(* IEC 61131-3 sources: daoli-st-library/DL_Device (part 42) *)

(* ---- FB_DL_PumpCavitationGuard.st ---- *)
(*==============================================================================
 * 组件名称 (Component)  : FB_DL_PumpCavitationGuard
 * 所属子库 (Sublibrary) : DL_Device
 * 当前版本 (Version)    : 1.0.1
 * 兼容性   (Platform)   : CODESYS 3.5 / TwinCAT 3 / 汇川 InoProShop / Schneider
 *                         Machine Expert；纯 IEC 61131-3（第 3 版）语法，
 *                         仅依赖 Standard.library（R_TRIG / TON）
 * 组件分类 (Category)   : 功能块（FUNCTION_BLOCK）· 设备本体退化诊断 · 泵汽蚀
 * 功能描述 (Function)   : 泵汽蚀的在线判据与**降速请求**。三判据并发：
 *                         (a) 流量偏低（低于额定的比例）；(b) 扬程跌落（低于额定的
 *                         跌幅）；(c) 振动超限**或**电流波动超限。三者同拍成立并
 *                         持续 tConfirm 才升级为锁存故障；单条成立只到「嫌疑」。
 * 降速语义 (Derate)     : 本件**不直接给变频器频率**，只输出 `fDerateRatio`
 *                         （1.0 = 不降）与 `bDerateRequest`。执行归上层
 *                         `FB_DL_RateLimiter` / `FB_DL_VfdGeneric`——诊断件一旦
 *                         自己写频率，就会与工艺主控的速率限制打架，且无法在
 *                         不同变频器之间移植。
 *                         每次确认汽蚀事件比率递减一步（下限 0.3），**只减不自动
 *                         增**：回升由上层斜坡完成，避免本件与上层同时调节同
 *                         一个量（双写冲突）。
 * 边界声明 (Limits)     : ① **不做 NPSH 计算**：需介质饱和蒸汽压与吸入侧压力，
 *                         属选型设计而非在线判据；② 振动阈值默认取 ISO 10816
 *                         C 区边界 4.5 mm/s（**公知阈值，引脚可改**），头注释
 *                         注明出处与「仅参考」定位；③ 本件**不声称**符合
 *                         ISO 10816 认证，阈值只是工程默认值；④ 停泵（bRunning
 *                         为 FALSE）时全部判据抑制，不产生任何降速请求。
 * 段序 (Cycle order)   : 段 1 默认值与单拍预清零 → 段 2 首扫初始化 →
 *                         段 3 参数闸门与输入域检查 → 段 4 定时器与边沿无条件刷新 →
 *                         段 5 判据计算 → 段 6 复位通道与故障锁存（**CASE 前置，
 *                         不做状态变量赋值**）→ 段 7 监视相位机 → 段 8 降速执行与
 *                         事件锁存 → 段 9 健康仲裁、出口钳位与保持重写 → 段 10 码位链。
 * 拍间依赖 (Cycle dep)  : 确认定时器在段 4 调用，而其 IN 里的「三判据同拍」在段 5
 *                         才算出，故定时器读到的是**上一拍照**的判据值（一拍滞后）。
 *                         对 3 秒量级的确认判据无实质影响，换来的是「所有定时器
 *                         实例都在同一段无条件调用」这一更强的纪律；此处显式登记，
 *                         避免后人误以为是笔误。
 * 定时器清单 (R40)      : 实例名 / IN 表达式 / 断输入拍标志 / 自清位置
 *                         fbConfirmWatch / 三判据同拍 AND 状态为嫌疑 AND
 *                                        NOT _bConfirmBreak / _bConfirmBreak
 *                                        （进/出嫌疑态与复位时置位）
 *                         fbRippleWatch  / 泵运行 AND NOT _bRippleBreak
 *                                        / _bRippleBreak（窗满后置位重启）
 *                         fbHoldOffWatch / 状态为降速 AND NOT _bHoldBreak
 *                                        / _bHoldBreak（进/出降速态置位）
 *                         三个实例全部在段 4 无条件调用，断输入拍一律在调用后自清。
 * 单拍标志清单 (R25)    : `_bResetPulse` 预清段 1 / 置位段 6 / 消费段 6；
 *                         `_bDerateStep`（降速单拍）预清段 1 / 置位段 8 / 消费段 8；
 *                         `_bConfirmEvent` 预清段 1 / 置位段 7 / 消费段 8；
 *                         三个断输入标志就地置位、段 4 调用后自清。
 * 保持位清单 (R27)      : `bDerateRequest` 与 `fDerateRatio`、`bCavitation`、
 *                         `nEventCount` 四个保持量，全部由段 9 每拍重写出口；
 *                         降速请求在 eDerate 与抑制窗内**保持为 TRUE**，不靠
 *                         进入那一拍的脉冲（R27 的典型场景）。
 * 三元一致表 (R35)      : 量 / 守卫封顶 / 判据运算符
 *                         fFlowLowRatio   / 钳到 0.2~0.95 / 判据用 <
 *                         fHeadDropRatio  / 钳到 0.05~0.5 / 判据用（1 减比值）>
 *                         fVibLimit       / 钳到 1~20     / 判据用比值 > 1，急停用 > 2
 *                         振动比值输出上限 / 钳到 5.0     / 必须高于急停倍率 2（R35 同向）
 *                         fDerateStep     / 钳到 0.02~0.3 / 递减后与 0.3 取大
 * 验收向量 (Acceptance) :
 *   V1 单判据：流量 0.5 倍额定（其余判据不成立）→ eSuspect + 0164，**不锁存**
 *   V2 三判据：三判据同拍持续 3 s → eConfirm → eDerate、0326、比率每次 −0.10
 *      （下限 0.3）
 *   V3（V-C 跨段 R40）：tConfirm 定时器在 eSuspect 与 eMonitor 来回时必须断输入，
 *      否则三次 1 s 的孤立嫌疑会被误判成「持续 3 s」
 *   V4（V-D 恢复）：bReset 后 fDerateRatio **不得**直接回 1.0（R41），且必须夹进
 *      0.3~1.0（R43）
 *   V5（V-A 域外）：fFlowNominal 为 0 → 0328 锁存，fFlowRatio 输出 0（不输出无穷大）
 * 规格偏离 (Deviation)  :
 *   ① 规格 V1 给的是「流量 0.5 倍额定、扬程 0.8 倍额定、振动 2.0、电流平稳 →
 *      只有流量判据」。按默认 fHeadDropRatio 为 0.15 计算，扬程 0.8 倍额定的跌幅
 *      为 20%，**会同时触发扬程判据**。本件按判据定义实现（跌幅 > 15% 即成立），
 *      复现 V1 需把 fHeadDropRatio 调到 ≥0.25；此处不改判据语义以迁就向量。
 *   ② 规格未给「电流波动率」的确切口径。本件取滑动窗内「(最大 − 最小) ÷ 平均」
 *      作为波动率，窗长 tRippleWindow，窗满即出值并重启窗；该口径与现场常见的
 *      「电流摆动幅度百分比」一致，且不依赖频谱。
 *   ③ 规格要求 bReset 后比率不直接回 1.0。本件在 bReset 且三判据全部消失时让
 *      比率**回升一步**（不直接回 1.0），其余恢复速率仍交上层斜坡；这是「不得
 *      重头恢复」与「不能让比率永久卡死」之间的折中，已在此登记。
 *   ④ 参数非法（额定值非正、阈值倒置）统一用 0328，未分更细码位（本轮未分配）。
 * 开源溯源 (Origin)     : 来源标签 namur-ne107 / lbp-basic-process / pump-diag。
 *                         原创 clean-room 实现。**仅借鉴**：① NAMUR NE107（公开
 *                         推荐规范）的健康分级语义；② LBP（Library of Basic
 *                         Process）公开文档所呈现的「命令—监视—判定」三段式
 *                         分层惯例，作为本件「判据—定级—降速请求」的组织参照。
 *                         汽蚀三判据（流量低 / 扬程跌 / 振动或电流波动）属泵
 *                         行业公开的通行定性认识；ISO 10816 的 4.5 mm/s 为公知
 *                         阈值。本件未复制任何源码行、未沿用其命名体系，窗口
 *                         口径、状态机、宽限与降速规则、全部码位 100% 本库独立
 *                         设计，无许可证传染风险。
 * 修订历史 (Revision)   :
 *   2026-11-15  v1.0.0  首版入库（R13 · 泳道 A · 泵汽蚀判据与降速请求）
 *   2026-11-16  v1.0.1  终审修复五处：① `_bHoldActive` 由「窗满那一拍」改为
 *                       「整个降速相」——原实现下 0165 仅在抑制窗到期瞬间可见、
 *                       判据在窗内并未被真正抑制；② 流量/扬程比值改用**原始
 *                       额定值的域**做门（原实现拿兜底值 1.0 当分母，额定为 0
 *                       时输出的是伪比值而非 0，违 V5）；③ 汽蚀确认补写
 *                       `_uErrFault := 16#0003_0326`（原实现 bError 为真而
 *                       uErrorId 恒 0，违 R21 一致性）；④ 急停级 0327 加
 *                       bRunning/bEnable 门（停泵时邻近设备振动不得拉锁存）；
 *                       ⑤ 停泵清 `_fRipple`，防停泵前旧波动率跨停机存活到
 *                       重启后的首个取样窗。
 *============================================================================*)

(*-----------------------------------------------------------------------------
 * 枚举: E_DL_CavitationState（归属本功能块，同文件发布）
 * 含义: 汽蚀监视相位。6 个成员在段 6 各有唯一标签，ELSE 只接脏值。
 *-----------------------------------------------------------------------------*)
TYPE E_DL_CavitationState :
(
    eIdle    := 0,     // 待机：未使能或停泵 / Idle, disabled or the pump is stopped
    eMonitor := 10,    // 监视：泵运行，判据全部不成立 / Monitoring, no criterion active
    eSuspect := 20,    // 嫌疑：单判据成立，未确认 / Suspect, one criterion active
    eConfirm := 30,    // 确认：三判据同拍且持续满足 / Confirm, all three held long enough
    eDerate  := 40,    // 降速：已请求降速，处于抑制窗 / Derate, request held during the hold-off
    eFault   := 99     // 故障：参数非法或振动急停级，锁存 / Fault, latched
);
END_TYPE

FUNCTION_BLOCK FB_DL_PumpCavitationGuard
VAR_INPUT
    bEnable             : BOOL;                      // 使能 [-] / Enable
    bReset              : BOOL;                      // 复位锁存，上升沿有效 [-] / Rising edge resets the latch
    bRunning            : BOOL;                      // 泵运行中，停泵时全部判据抑制 [-] / Pump running, criteria suppressed when stopped
    fFlow               : REAL;                      // 实测流量 [m³/h]，范围 0~100000 / Measured flow
    fHead               : REAL;                      // 实测扬程 [m]，范围 0~1000 / Measured head
    fVibration          : REAL;                      // 振动速度有效值 [mm/s]，范围 0~50 / Vibration RMS velocity
    fCurrent            : REAL;                      // 电机电流 [A]，范围 0~10000 / Motor current
    fFlowNominal        : REAL;                      // 额定流量 [m³/h]，域大于 0 / Nominal flow, must exceed zero
    fHeadNominal        : REAL;                      // 额定扬程 [m]，域大于 0 / Nominal head, must exceed zero
    fFlowLowRatio       : REAL := 0.60;              // 流量低于额定的比例 [-]，范围 0.2~0.95 / Low-flow ratio
    fHeadDropRatio      : REAL := 0.15;              // 扬程跌落比例 [-]，范围 0.05~0.5 / Head-drop ratio
    fVibLimit           : REAL := 4.5;               // 振动上限 [mm/s]，ISO 10816 C 区边界，范围 1~20 / Vibration limit
    fCurrentRippleLimit : REAL := 0.15;              // 电流波动率上限 [-]，范围 0.02~0.5 / Current ripple limit
    tRippleWindow       : TIME := T#2S;              // 电流波动统计窗 [毫秒]，范围 0.5~30 s / Ripple window
    tConfirm            : TIME := T#3S;              // 三判据同拍持续判据 [毫秒]，范围 0.5~30 s / Confirmation time
    tHoldOff            : TIME := T#30S;             // 降速后抑制判据时长 [毫秒]，范围 5 s~10 min / Hold-off after a derate
    fDerateStep         : REAL := 0.10;              // 每次降速步长 [-]，范围 0.02~0.3 / Derate step
END_VAR
VAR_OUTPUT
    eHealth             : E_DL_Ne107Status;          // NE107 健康态（引用自 I_DL_DeviceHealth）[-] / NE107 health
    uDiagCode           : UDINT;                     // 当前诊断码，0=无码 [代码] / Active diagnostic code
    uErrorId            : UDINT;                     // 末次故障码，仅故障级 [代码] / Last fault code
    bError              : BOOL;                      // 故障锁存 [-] / Fault latched
    bCavitation         : BOOL;                      // 汽蚀确认（三判据同拍成立，锁存）[-] / Cavitation confirmed, latched
    bDerateRequest      : BOOL;                      // 降速请求（保持语义）[-] / Derate request, held
    fDerateRatio        : REAL;                      // 降速比例 [-]，范围 0.3~1.0，1.0=不降 / Derate ratio
    fFlowRatio          : REAL;                      // 实测/额定流量比值 [-]，钳 0~2 / Flow ratio
    fHeadRatio          : REAL;                      // 实测/额定扬程比值 [-]，钳 0~2 / Head ratio
    fVibRatio           : REAL;                      // 振动/上限比值 [-] / Vibration ratio
    nEventCount         : UDINT;                     // 汽蚀事件累计 [次]，锁存 / Event counter
    fRippleMeas         : REAL;                      // 窗内电流波动率实测值 [-] / Measured ripple
END_VAR
VAR
    fbTrigReset     : R_TRIG;                        // 复位沿检测，段 4 无条件刷新 [-] / Reset edge detector
    fbConfirmWatch  : TON;                           // 三判据持续计时，段 4 刷新 [毫秒] / Confirmation timer
    fbRippleWatch   : TON;                           // 电流波动统计窗，段 4 刷新 [毫秒] / Ripple window timer
    fbHoldOffWatch  : TON;                           // 降速后抑制窗，段 4 刷新 [毫秒] / Hold-off timer
    _eState         : E_DL_CavitationState := E_DL_CavitationState.eIdle; // 当前相位 [-] / Current phase
    _bInit          : BOOL := FALSE;                 // 首扫标志，初值 FALSE [-] / First-scan flag
    _bFaultLatch    : BOOL;                          // 故障锁存，仅复位清 [-] / Fault latch
    _uErrFault      : UDINT;                         // 首出故障码 [代码] / First-out fault code
    _uDiagCode      : UDINT;                         // 当前诊断码（单一链产出）[代码] / Active diagnostic code
    _bResetPulse    : BOOL;                          // 复位单拍 [-] / One-shot reset
    _bParamBad      : BOOL;                          // 参数非法标志 [-] / Illegal parameter flag
    _bConfirmBreak  : BOOL;                          // 确认定时器断输入一拍 [-] / Confirmation timer break
    _bRippleBreak   : BOOL;                          // 波动窗断输入一拍 [-] / Ripple window break
    _bHoldBreak     : BOOL;                          // 抑制窗断输入一拍 [-] / Hold-off break
    _fFlowNomUse    : REAL := 1.0;                   // 生效额定流量 [m³/h] / Effective nominal flow
    _fHeadNomUse    : REAL := 1.0;                   // 生效额定扬程 [m] / Effective nominal head
    _fFlowLowUse    : REAL := 0.60;                  // 生效流量比例 [-] / Effective low-flow ratio
    _fHeadDropUse   : REAL := 0.15;                  // 生效扬程跌幅 [-] / Effective head-drop ratio
    _fVibUse        : REAL := 4.5;                   // 生效振动上限 [mm/s] / Effective vibration limit
    _fRippleLimUse  : REAL := 0.15;                  // 生效波动率上限 [-] / Effective ripple limit
    _fStepUse       : REAL := 0.10;                  // 生效降速步长 [-] / Effective derate step
    _tRippleUse     : TIME := T#2S;                  // 生效波动窗 [毫秒] / Effective ripple window
    _tConfirmUse    : TIME := T#3S;                  // 生效确认时长 [毫秒] / Effective confirmation time
    _tHoldUse       : TIME := T#30S;                 // 生效抑制窗 [毫秒] / Effective hold-off
    _diMs           : DINT;                          // 时间换算中间量 [毫秒] / Time conversion working value
    _fFlowRatio     : REAL;                          // 流量比值 [-]，钳 0~2 / Flow ratio
    _fHeadRatio     : REAL;                          // 扬程比值 [-]，钳 0~2 / Head ratio
    _fVibRatio      : REAL;                          // 振动比值 [-] / Vibration ratio
    _bCritFlow      : BOOL;                          // 流量判据 [-] / Flow criterion
    _bCritHead      : BOOL;                          // 扬程判据 [-] / Head criterion
    _bCritVib       : BOOL;                          // 振动判据 [-] / Vibration criterion
    _bCritRipple    : BOOL;                          // 电流波动判据 [-] / Ripple criterion
    _bCritVibGroup  : BOOL;                          // 振动或波动（第三判据）[-] / Vibration or ripple, the third criterion
    _bAllThree      : BOOL;                          // 三判据同拍成立 [-] / All three criteria in one scan
    _bAnyCrit       : BOOL;                          // 任一判据成立 [-] / Any criterion active
    _bVibEmergency  : BOOL;                          // 振动超上限两倍（急停级）[-] / Vibration above twice the limit
    _fCurrMin       : REAL;                          // 窗内电流最小值 [A] / Minimum current in the window
    _fCurrMax       : REAL;                          // 窗内电流最大值 [A] / Maximum current in the window
    _fCurrSum       : REAL;                          // 窗内电流累加 [A] / Current sum in the window
    _nCurrCount     : UDINT;                         // 窗内电流样本数 [个] / Current sample count
    _fRipple        : REAL;                          // 窗内波动率实测值 [-] / Measured ripple
    _bHoldActive    : BOOL;                          // 抑制窗生效中 [-] / Hold-off active
    _bDerateStep    : BOOL;                          // 本次确认需降一步 [-] / Step down this scan
    _bConfirmEvent  : BOOL;                          // 本拍确认事件 [-] / Confirmation event this scan
    _bCavLatch      : BOOL;                          // 汽蚀锁存 [-] / Cavitation latch
    _fDerateRatio   : REAL := 1.0;                   // 保持的降速比例 [-] / Held derate ratio
    _bDerateHeld    : BOOL;                          // 保持的降速请求 [-] / Held derate request
    _uEventCount    : UDINT;                         // 保持的事件计数 [次] / Held event counter
    _eHealthInt     : E_DL_Ne107Status := E_DL_Ne107Status.eUnknown; // 健康态内部量 [-] / Internal health state
END_VAR
VAR CONSTANT
    DL_VAL_LIM      : REAL := 1.0E6;                 // 有限性判定绝对值上限 [-] / Finiteness limit
    DL_EPS          : REAL := 1.0E-6;                // 浮点比较容差 [-] / Float comparison tolerance
    DL_RATIO_MAX    : REAL := 2.0;                   // 流量扬程比值上限 [-]，防噪声放大 / Flow and head ratio ceiling
    DL_VIB_RATIO_MAX: REAL := 5.0;                   // 振动比值上限 [-]，须高于急停倍率 2 倍（R35 同向） / Vibration ratio ceiling
    DL_VIB_EMERG    : REAL := 2.0;                   // 振动急停级倍率 [-] / Emergency vibration multiplier
    DL_DERATE_MIN   : REAL := 0.3;                   // 降速比例下限 [-] / Lower derate bound
    DL_DERATE_MAX   : REAL := 1.0;                   // 降速比例上限 [-] / Upper derate bound
    DL_RIPPLE_MIN_MS: DINT := 500;                   // 波动窗下限 [毫秒] / Minimum ripple window
    DL_RIPPLE_MAX_MS: DINT := 30000;                 // 波动窗上限 [毫秒] / Maximum ripple window
    DL_CONFIRM_MIN  : DINT := 500;                   // 确认时长下限 [毫秒] / Minimum confirmation
    DL_CONFIRM_MAX  : DINT := 30000;                 // 确认时长上限 [毫秒] / Maximum confirmation
    DL_HOLD_MIN     : DINT := 5000;                  // 抑制窗下限 [毫秒] / Minimum hold-off
    DL_HOLD_MAX     : DINT := 600000;                // 抑制窗上限 [毫秒] / Maximum hold-off
END_VAR

(*------------------------------------------------------------------------------
 * 段 1｜确定性默认值与单拍标志预清零（R25 第一律）
 *      Deterministic defaults and one-shot flags pre-cleared
 *-----------------------------------------------------------------------------*)
_bResetPulse   := FALSE;                              // 复位单拍预清零（Reset pre-cleared）
_bParamBad     := FALSE;                              // 参数非法预清零（Illegal parameter pre-cleared）
_bDerateStep   := FALSE;                              // 降速单拍预清零（Derate step pre-cleared）
_bConfirmEvent := FALSE;                              // 确认事件预清零（Confirmation event pre-cleared）
_bCritFlow     := FALSE;                              // 流量判据预清零（Flow criterion pre-cleared）
_bCritHead     := FALSE;                              // 扬程判据预清零（Head criterion pre-cleared）
_bCritVib      := FALSE;                              // 振动判据预清零（Vibration criterion pre-cleared）
_bCritRipple   := FALSE;                              // 波动判据预清零（Ripple criterion pre-cleared）
_bVibEmergency := FALSE;                              // 振动急停预清零（Emergency pre-cleared）

(*------------------------------------------------------------------------------
 * 段 2｜首扫初始化（R19：bInit 初值 FALSE，判据取非；首拍只装基准）
 *      First-scan initialisation, baseline only
 *-----------------------------------------------------------------------------*)
IF NOT _bInit THEN
    _eState       := E_DL_CavitationState.eIdle;      // 相位待机（Phase idle）
    _bFaultLatch  := FALSE;                           // 故障锁存清零（Latch cleared）
    _uErrFault    := 16#0000_0000;                    // 首出码清零（First-out code cleared）
    _bCavLatch    := FALSE;                           // 汽蚀锁存清零（Cavitation latch cleared）
    _fDerateRatio := DL_DERATE_MAX;                   // 冷启动比率 1.0，落在有效域内（Cold start at 1.0）
    _bDerateHeld  := FALSE;                           // 降速请求清零（Derate request cleared）
    _uEventCount  := 0;                               // 事件计数清零（Event counter cleared）
    _fRipple      := 0.0;                             // 波动率初值 0（Ripple starts at zero）
    _fCurrMin     := DL_VAL_LIM;                      // 最小值先置上界（Minimum preset to the ceiling）
    _fCurrMax     := 0.0;                             // 最大值先置 0（Maximum preset to zero）
    _fCurrSum     := 0.0;                             // 电流累加清零（Current sum cleared）
    _nCurrCount   := 0;                               // 样本数清零（Sample count cleared）
    _fFlowNomUse  := 1.0;                             // 额定流量兜底（Nominal flow fallback）
    _fHeadNomUse  := 1.0;                             // 额定扬程兜底（Nominal head fallback）
    _bInit        := TRUE;                            // 首扫只做一次（First scan runs once）
END_IF

(*------------------------------------------------------------------------------
 * 段 3｜参数闸门与输入域检查（额定值非正或阈值倒置属故障级）
 *      Parameter gate: non-positive nominals or inverted thresholds latch a fault
 *-----------------------------------------------------------------------------*)
IF (fFlowNominal <= DL_EPS) OR (fHeadNominal <= DL_EPS) OR (fVibLimit <= DL_EPS) THEN
    _bParamBad := TRUE;                               // 额定值或振动上限非正（Non-positive nominals）
END_IF
IF (fFlowLowRatio <= 0.0) OR (fFlowLowRatio >= 1.0) OR (fHeadDropRatio <= 0.0) OR (fHeadDropRatio >= 1.0) THEN
    _bParamBad := TRUE;                               // 比例阈值倒置（Inverted ratios）
END_IF
IF (fCurrentRippleLimit <= 0.0) OR (fDerateStep <= 0.0) OR (fDerateStep > 0.5) THEN
    _bParamBad := TRUE;                               // 波动限或步长非法（Illegal ripple limit or step）
END_IF

IF fFlowNominal > DL_EPS THEN
    _fFlowNomUse := fFlowNominal;                     // 额定流量直通（Nominal flow passed through）
ELSE
    _fFlowNomUse := 1.0;                              // 非正：兜底为 1，防除零（Fallback avoids a zero divisor）
END_IF
IF fHeadNominal > DL_EPS THEN
    _fHeadNomUse := fHeadNominal;                     // 额定扬程直通（Nominal head passed through）
ELSE
    _fHeadNomUse := 1.0;                              // 非正：兜底为 1（Fallback）
END_IF

_fFlowLowUse   := LIMIT(0.2, fFlowLowRatio, 0.95);    // 流量比例钳进 0.2~0.95（Clamped）
_fHeadDropUse  := LIMIT(0.05, fHeadDropRatio, 0.5);   // 跌幅比例钳进 0.05~0.5（Clamped）
_fVibUse       := LIMIT(1.0, fVibLimit, 20.0);        // 振动上限钳进 1~20 mm/s（Clamped）
_fRippleLimUse := LIMIT(0.02, fCurrentRippleLimit, 0.5); // 波动限钳进 0.02~0.5（Clamped）
_fStepUse      := LIMIT(0.02, fDerateStep, 0.3);      // 降速步长钳进 0.02~0.3（Clamped）

_diMs         := LIMIT(DL_RIPPLE_MIN_MS, TIME_TO_DINT(tRippleWindow), DL_RIPPLE_MAX_MS); // 波动窗钳位（Clamped）
_tRippleUse   := DINT_TO_TIME(_diMs);                 // 生效波动窗（Effective ripple window）
_diMs         := LIMIT(DL_CONFIRM_MIN, TIME_TO_DINT(tConfirm), DL_CONFIRM_MAX); // 确认时长钳位（Clamped）
_tConfirmUse  := DINT_TO_TIME(_diMs);                 // 生效确认时长（Effective confirmation）
_diMs         := LIMIT(DL_HOLD_MIN, TIME_TO_DINT(tHoldOff), DL_HOLD_MAX); // 抑制窗钳位（Clamped）
_tHoldUse     := DINT_TO_TIME(_diMs);                 // 生效抑制窗（Effective hold-off）

(*------------------------------------------------------------------------------
 * 段 4｜定时器与边沿实例无条件刷新（红线：实例一律在 CASE 之外每拍必调）
 *      Timers and edge detectors refreshed unconditionally outside the CASE
 *-----------------------------------------------------------------------------*)
fbTrigReset(CLK := bReset);                           // 复位沿刷新（Reset edge refreshed）

fbConfirmWatch(IN := _bAllThree AND (_eState = E_DL_CavitationState.eSuspect) AND (NOT _bConfirmBreak), PT := _tConfirmUse); // 三判据持续计时
_bConfirmBreak := FALSE;                              // 断输入拍在调用后自清（Break self-cleared）

fbRippleWatch(IN := bRunning AND (NOT _bRippleBreak), PT := _tRippleUse); // 波动统计窗
_bRippleBreak := FALSE;                               // 断输入拍在调用后自清（Break self-cleared）

fbHoldOffWatch(IN := (_eState = E_DL_CavitationState.eDerate) AND (NOT _bHoldBreak), PT := _tHoldUse); // 抑制窗计时
_bHoldBreak := FALSE;                                 // 断输入拍在调用后自清（Break self-cleared）
_bHoldActive := (_eState = E_DL_CavitationState.eDerate) OR fbHoldOffWatch.Q; // 抑制生效 = 整个降速相（不是窗满那一拍）

(*------------------------------------------------------------------------------
 * 段 5｜判据计算（比值前置守卫，绝不输出无穷大；V5）
 *      Criteria, ratios guarded against division by zero
 *-----------------------------------------------------------------------------*)
(* 比值口径：额定值非正时**输出 0**，绝不拿兜底值 1.0 去算伪比值（V5 明确要求） *)
IF fFlowNominal > DL_EPS THEN
    _fFlowRatio := LIMIT(0.0, fFlow / _fFlowNomUse, DL_RATIO_MAX); // 流量比值，钳 0~2（Clamped）
ELSE
    _fFlowRatio := 0.0;                               // 额定流量非法：输出 0，不给伪比值（Never a pseudo ratio）
END_IF
IF fHeadNominal > DL_EPS THEN
    _fHeadRatio := LIMIT(0.0, fHead / _fHeadNomUse, DL_RATIO_MAX); // 扬程比值，钳 0~2（Clamped）
ELSE
    _fHeadRatio := 0.0;                               // 额定扬程非法：输出 0（Never a pseudo ratio）
END_IF
IF _fVibUse > DL_EPS THEN
    _fVibRatio := LIMIT(0.0, fVibration / _fVibUse, DL_VIB_RATIO_MAX); // 振动比值，上限须容得下急停倍率（Clamped）
ELSE
    _fVibRatio := 0.0;                                // 分母不可用：输出 0（Never infinity）
END_IF

(* 三判据：停泵或抑制窗内一律不成立（Suppressed when stopped or within the hold-off） *)
IF bRunning AND bEnable AND (NOT _bHoldActive) THEN
    _bCritFlow   := _fFlowRatio < _fFlowLowUse;                       // 流量偏低（Low flow）
    _bCritHead   := _fHeadRatio < (1.0 - _fHeadDropUse);              // 扬程跌落（Head drop）
    _bCritVib    := _fVibRatio > 1.0;                                 // 振动超限（Vibration above limit）
    _bCritRipple := _fRipple > _fRippleLimUse;                        // 电流波动超限（Ripple above limit）
END_IF
_bCritVibGroup := _bCritVib OR _bCritRipple;                          // 第三判据：振动或波动（Third criterion）
_bAllThree     := _bCritFlow AND _bCritHead AND _bCritVibGroup;       // 三判据同拍（All three in one scan）
_bAnyCrit      := _bCritFlow OR _bCritHead OR _bCritVibGroup;         // 任一判据（Any criterion）
(* 急停级：仅在泵运行且使能时成立。停泵时邻近设备振动/传感器卡值不得把本件拉进锁存，
 * 与「bRunning 为 FALSE 时全部判据抑制」同一条纪律；降速抑制窗内仍照判（等级高于判据） *)
IF bRunning AND bEnable AND (_fVibRatio > DL_VIB_EMERG) THEN
    _bVibEmergency := TRUE;                                           // 振动超两倍上限（Emergency level）
END_IF

(* 电流波动统计：窗满出一值并重启窗（Window closes, one value produced, window restarts） *)
IF bRunning THEN
    IF fCurrent < _fCurrMin THEN
        _fCurrMin := fCurrent;                        // 更新最小（Update the minimum）
    END_IF
    IF fCurrent > _fCurrMax THEN
        _fCurrMax := fCurrent;                        // 更新最大（Update the maximum）
    END_IF
    _fCurrSum := _fCurrSum + fCurrent;                // 累加（Accumulate）
    IF _nCurrCount < 16#FFFF_FFFF THEN
        _nCurrCount := _nCurrCount + 1;               // 计数防上溢（Guard the counter）
    END_IF
    IF fbRippleWatch.Q THEN
        IF _nCurrCount > 0 THEN
            IF (_fCurrSum / UDINT_TO_REAL(_nCurrCount)) > DL_EPS THEN
                _fRipple := (_fCurrMax - _fCurrMin) / (_fCurrSum / UDINT_TO_REAL(_nCurrCount)); // 波动率，分母已守卫
            ELSE
                _fRipple := 0.0;                      // 平均近零：不判波动（No meaningful ripple）
            END_IF
        END_IF
        _fCurrMin   := DL_VAL_LIM;                    // 窗重启：最小值复位（Window restarted）
        _fCurrMax   := 0.0;                           // 窗重启：最大值复位（Window restarted）
        _fCurrSum   := 0.0;                           // 窗重启：累加清零（Window restarted）
        _nCurrCount := 0;                             // 窗重启：计数清零（Window restarted）
        _bRippleBreak := TRUE;                        // 断输入一拍后重新计时（One-scan break restarts the timer）
    END_IF
ELSE
    _fCurrMin   := DL_VAL_LIM;                        // 停泵清零（Cleared while stopped）
    _fCurrMax   := 0.0;                               // 停泵清零（Cleared while stopped）
    _fCurrSum   := 0.0;                               // 停泵清零（Cleared while stopped）
    _nCurrCount := 0;                                 // 停泵清零（Cleared while stopped）
    _fRipple    := 0.0;                               // 停泵清实测值，防停泵前旧值跨停机存活（Stale ripple must not survive a stop）
END_IF

(*------------------------------------------------------------------------------
 * 段 6｜复位通道 + 故障锁存（CASE 前置；**不做状态变量赋值**，R39）
 *      Reset channel and fault latching before the CASE, with no state write
 *-----------------------------------------------------------------------------*)
IF fbTrigReset.Q THEN
    _bResetPulse := TRUE;                             // 复位单拍（One-shot reset）
END_IF

IF _bResetPulse THEN
    _bFaultLatch := FALSE;                            // 清故障锁存（Latch cleared）
    _uErrFault   := 16#0000_0000;                     // 清首出码（First-out code cleared）
    _bCavLatch   := FALSE;                            // 清汽蚀锁存（Cavitation latch cleared）
    _bDerateHeld := FALSE;                            // 撤降速请求，交给上层斜坡（Release the request to the upper ramp）
    IF _bAnyCrit THEN
        _fDerateRatio := LIMIT(DL_DERATE_MIN, _fDerateRatio, DL_DERATE_MAX); // 判据仍在：比率保持并夹域（Held while criteria persist）
    ELSE
        _fDerateRatio := LIMIT(DL_DERATE_MIN, _fDerateRatio + _fStepUse, DL_DERATE_MAX); // 判据已消：回升一步，不直接回 1.0（R41）
    END_IF
    _bConfirmBreak := TRUE;                           // 确认计时重启（Confirmation timer restarted）
    _bRippleBreak  := TRUE;                           // 波动窗重启（Ripple window restarted）
    _bHoldBreak    := TRUE;                           // 抑制窗重启（Hold-off restarted）
END_IF

IF _bParamBad AND (NOT _bFaultLatch) THEN
    _uErrFault   := 16#0003_0328;                     // 0328 额定值非正或阈值倒置（Illegal nominals or thresholds）
    _bFaultLatch := TRUE;                             // 锁存（Latched）
END_IF

(*------------------------------------------------------------------------------
 * 段 7｜监视相位机（6 个成员各一标签 + ELSE 兜底）
 *      Monitoring state machine, one label per member plus a trailing fallback
 *-----------------------------------------------------------------------------*)
CASE _eState OF

    E_DL_CavitationState.eIdle: // 待机：起泵后进入监视
        IF _bFaultLatch THEN
            _eState := E_DL_CavitationState.eFault;   // 已锁故障（Already latched）
        ELSIF bEnable AND bRunning THEN
            _bConfirmBreak := TRUE;                   // 确认计时从 0 起算（Confirmation restarts）
            _bRippleBreak  := TRUE;                   // 波动窗从 0 起算（Ripple window restarts）
            _bHoldBreak    := TRUE;                   // 抑制窗从 0 起算（Hold-off restarts）
            _eState := E_DL_CavitationState.eMonitor; // 进监视（Enter monitoring）
        END_IF

    E_DL_CavitationState.eMonitor: // 监视：任一判据即进嫌疑
        IF _bFaultLatch THEN
            _eState := E_DL_CavitationState.eFault;   // 转故障（Enter the fault state）
        ELSIF (NOT bEnable) OR (NOT bRunning) THEN
            _eState := E_DL_CavitationState.eIdle;    // 停泵或掉使能回待机（Stopped or disabled, back to idle）
        ELSIF _bAnyCrit AND (NOT _bHoldActive) THEN
            _bConfirmBreak := TRUE;                   // 进嫌疑：确认计时从 0 起算（R40 段边界断输入）
            _eState := E_DL_CavitationState.eSuspect; // 进嫌疑（Enter suspect）
        END_IF

    E_DL_CavitationState.eSuspect: // 嫌疑：三判据同拍并持续满足才确认
        IF _bFaultLatch THEN
            _eState := E_DL_CavitationState.eFault;   // 转故障（Enter the fault state）
        ELSIF (NOT bEnable) OR (NOT bRunning) THEN
            _eState := E_DL_CavitationState.eIdle;    // 停泵回待机（Stopped, back to idle）
        ELSIF NOT _bAnyCrit THEN
            _bConfirmBreak := TRUE;                   // 判据消失：确认计时断输入（Criterion cleared, timer broken）
            _eState := E_DL_CavitationState.eMonitor; // 回监视（Back to monitoring）
        ELSIF fbConfirmWatch.Q THEN
            _bConfirmEvent := TRUE;                   // 确认事件单拍（Confirmation event）
            _eState := E_DL_CavitationState.eConfirm; // 进确认（Enter confirmation）
        END_IF

    E_DL_CavitationState.eConfirm: // 确认：本拍锁存并请求降速，随后进入降速相
        _bConfirmBreak := TRUE;                       // 确认计时清零（Confirmation cleared）
        _bHoldBreak    := TRUE;                       // 抑制窗从 0 起算（Hold-off restarts）
        _eState := E_DL_CavitationState.eDerate;      // 进降速（Enter derate）
        IF (NOT bEnable) OR (NOT bRunning) THEN
            _eState := E_DL_CavitationState.eIdle;    // 停泵中止（Stopped, abort）
        END_IF

    E_DL_CavitationState.eDerate: // 降速：抑制窗内忽略判据，窗满且判据消失才回监视
        IF _bFaultLatch THEN
            _eState := E_DL_CavitationState.eFault;   // 转故障（Enter the fault state）
        ELSIF (NOT bEnable) OR (NOT bRunning) THEN
            _bHoldBreak := TRUE;                      // 抑制窗中断（Hold-off stopped）
            _eState := E_DL_CavitationState.eIdle;    // 停泵回待机（Stopped, back to idle）
        ELSIF fbHoldOffWatch.Q THEN
            (* 抑制窗内判据被强制为假，故出口条件只看窗满；窗满后判据在
             * eMonitor 重新评估，若仍成立会再次进入嫌疑并再降一步 *)
            _bHoldBreak := TRUE;                      // 抑制窗结束重启（Hold-off finished）
            _bDerateHeld := FALSE;                    // 撤降速请求，交由上层斜坡（Request released to the upper ramp）
            _bConfirmBreak := TRUE;                   // 确认计时重启（Confirmation restarted）
            _eState := E_DL_CavitationState.eMonitor; // 回监视（Back to monitoring）
        END_IF

    E_DL_CavitationState.eFault: // 故障：等复位
        IF _bResetPulse THEN
            _eState := E_DL_CavitationState.eIdle;    // 复位受理（Reset accepted）
        END_IF

    ELSE
        _uErrFault   := 16#0003_0329;                 // 0329 非法状态兜底（Illegal state fallback）
        _bFaultLatch := TRUE;                         // 兜底锁存（Fallback latched）
        _eState      := E_DL_CavitationState.eFault;  // 进终端安全态（Terminal safe state）
END_CASE

(*------------------------------------------------------------------------------
 * 段 8｜降速执行与事件锁存（确认事件、步进、急停级）
 *      Derate execution and event latching
 *-----------------------------------------------------------------------------*)
IF _bConfirmEvent THEN
    _bCavLatch := TRUE;                               // 汽蚀锁存（Cavitation latched）
    IF NOT _bFaultLatch THEN
        _uErrFault := 16#0003_0326;                   // 汽蚀确认亦属故障级：写入末次故障码，防 bError 为真而 uErrorId 为 0（R21 一致性）
    END_IF
    _bDerateHeld := TRUE;                             // 降速请求保持（Request held）
    _bDerateStep := TRUE;                             // 本拍降一步（Step down this scan）
    IF _uEventCount < 16#FFFF_FFFF THEN
        _uEventCount := _uEventCount + 1;             // 事件计数（Event counter incremented）
    END_IF
    _bConfirmEvent := FALSE;                          // 单拍消费后自清（Event consumed）
END_IF

IF _bDerateStep THEN
    _fDerateRatio := LIMIT(DL_DERATE_MIN, _fDerateRatio - _fStepUse, DL_DERATE_MAX); // 递减一步并夹域（Step down, clamped）
    _bDerateStep := FALSE;                            // 单拍消费后自清（Step consumed）
END_IF

IF _bVibEmergency AND (NOT _bFaultLatch) THEN
    _uErrFault   := 16#0003_0327;                     // 0327 振动超两倍上限（Emergency vibration）
    _bFaultLatch := TRUE;                             // 锁存（Latched）
    _bCavLatch   := TRUE;                             // 急停级同样置汽蚀（Treated as cavitation evidence）
END_IF

IF (_eState = E_DL_CavitationState.eDerate) OR _bFaultLatch THEN
    _bDerateHeld := TRUE;                             // 降速态与故障态内请求保持（Request held in derate and fault）
END_IF

(*------------------------------------------------------------------------------
 * 段 9｜健康仲裁、出口钳位与保持重写（R27 + R43）
 *      Health arbitration, clamping and hold semantics
 *-----------------------------------------------------------------------------*)
IF _bFaultLatch OR _bCavLatch THEN
    _eHealthInt := E_DL_Ne107Status.eFailure;         // 失效：含汽蚀确认（Failure, including confirmed cavitation）
ELSIF _eState = E_DL_CavitationState.eSuspect THEN
    _eHealthInt := E_DL_Ne107Status.eOutOfSpec;       // 嫌疑：超出规格但未确认（Suspect, out of specification）
ELSIF NOT bEnable THEN
    _eHealthInt := E_DL_Ne107Status.eUnknown;         // 未使能（Disabled）
ELSE
    _eHealthInt := E_DL_Ne107Status.eOk;              // 正常（OK）
END_IF

eHealth        := _eHealthInt;                        // 健康态出口（Health outlet）
bCavitation    := _bCavLatch;                         // 汽蚀锁存保持重写（Held cavitation flag）
bDerateRequest := _bDerateHeld;                       // 降速请求保持重写（Held request rewritten）
fDerateRatio   := LIMIT(DL_DERATE_MIN, _fDerateRatio, DL_DERATE_MAX); // 比率钳进 0.3~1.0（Clamped, R43）
fFlowRatio     := LIMIT(0.0, _fFlowRatio, DL_RATIO_MAX); // 流量比值钳位（Clamped）
fHeadRatio     := LIMIT(0.0, _fHeadRatio, DL_RATIO_MAX); // 扬程比值钳位（Clamped）
fVibRatio      := LIMIT(0.0, _fVibRatio, DL_VIB_RATIO_MAX); // 振动比值钳位（Clamped）
nEventCount    := _uEventCount;                       // 事件计数出口（Event counter outlet）
fRippleMeas    := LIMIT(0.0, _fRipple, 10.0);          // 波动率出口钳进 0~10（Clamped）
bError         := _bFaultLatch OR _bCavLatch;          // 汽蚀确认亦属失效级（Confirmed cavitation is a failure）

(*------------------------------------------------------------------------------
 * 段 10｜码位单一优先级链（全拍只写一次 uDiagCode）
 *      Single priority chain, the diagnostic code is written exactly once
 *-----------------------------------------------------------------------------*)
IF _bFaultLatch THEN
    _uDiagCode := _uErrFault;                         // 故障级优先，保留首出码（Fault level, first-out code）
ELSIF _bCavLatch THEN
    _uDiagCode := 16#0003_0326;                       // 0326 汽蚀确认（Cavitation confirmed）
ELSIF (_eState = E_DL_CavitationState.eSuspect) THEN
    _uDiagCode := 16#0003_0164;                       // 0164 单判据嫌疑（Single criterion, suspect only）
ELSIF _bHoldActive THEN
    _uDiagCode := 16#0003_0165;                       // 0165 抑制窗内判据被忽略（Criteria ignored in the hold-off）
ELSE
    _uDiagCode := 16#0000_0000;                       // 无码（No code）
END_IF

uDiagCode := _uDiagCode;                              // 诊断码出口（Diagnostic code outlet）
uErrorId  := _uErrFault;                              // 末次故障码出口（Last fault code outlet）

END_FUNCTION_BLOCK

(* ---- FB_DL_RfidTagHandler.st ---- *)
(*==============================================================================
 * 组件名称 (Component)  : FB_DL_RfidTagHandler
 * 所属子库 (Sublibrary) : DL_Device
 * 当前版本 (Version)    : 1.0.1
 * 组件分类 (Category)   : 功能块（FUNCTION_BLOCK）· 设备实现件 · 状态机
 * 兼容性   (Platform)   : CODESYS 3.5 / TwinCAT 3 / 汇川 InoProShop / Schneider
 *                         Machine Expert；仅 Standard.library 的 TON 与 R_TRIG
 * 功能描述 (Function)   : I_DL_RfidReader 的标准实现件。以「请求 到 执行 到
 *                         应答」三拍握手驱动外部读写头（硬件经引脚注入就绪、
 *                         完成、报错、标签号、数据区、原始错误码，零硬编码
 *                         地址），内置单指令互斥、超时转重试转耗尽报错链、
 *                         同标签重复读抑制窗、写后回读校验、读写计数与诊断。
 * 双类故障 (Fault split) : 借 AOI 的「组态类与工艺类故障分离」思想，本块把
 *                         故障分两段：
 *                         组态与使用类 16#0003_02F0 / 02F1（忙时重入、写入内容
 *                         非法、超时重试耗尽）表示参数或调用方式有问题，
 *                         HMI 应提示改组态或查线缆；
 *                         工艺类 16#0003_02F2 / 02F3（读写头报错重试耗尽、
 *                         写后回读不符、非法状态兜底）表示硬件或工件有问题，
 *                         HMI 应提示叫维修。
 *                         两类同置 bError，但码段分开，便于报警分级。
 * 设计要点 (Key notes)  : ① 单指令互斥：忙态再调用读写方法一律返回 FALSE 并
 *                           置 02F0，不排队（硬件本身互斥，排队会让上层误判）；
 *                         ② 无标签是业务态（bNoTag）不是故障：不置 bError、
 *                           不计重试次数，HMI 直接提示「请放标签」；
 *                         ③ 计时器栅极复位范式：TON 复位只能靠 IN 拉低一整拍，
 *                           故用「栅极加再武装」两个标志实现，禁止用清 ET 的
 *                           厂商写法（ET 不可写才是跨平台共识）；
 *                         ④ 阈值三源优先级写死：常量域（最终兜底）低于引脚，
 *                           引脚低于 Init 注入的组态；同一字段只有一个方向，
 *                           不出现隐式切换；
 *                         ⑤ 单拍输出（bReadDoneOk / bWriteDoneOk）在主体首行
 *                           预清零（R25 律①）；bNoTag 与 Tag 快照为保持型
 *                           （R27），直到下一次成功或新指令开始。
 * 开源溯源 (Origin)     : tcopen-component / rockwell-aoi。参考 TcOpen 公开组件
 *                         库的契约实现分离与状态只读属性思想，以及 Rockwell AOI
 *                         公开手册所述参数分段与「程序类故障与操作类故障分离」
 *                         的组织方式。仅借组织思想与分类，状态机、码位、结构体
 *                         布局 100% 自有 clean-room，不构成衍生作品。
 * 依赖     (Depends)    : I_DL_RfidReader（本文件实现其全部 7 个成员）
 * 故障码表 (Error codes):
 *   16#0003_0138【信息级】同标签重复读被抑制窗拦下
 *   16#0003_0139【信息级】指令超时或抑制窗参数越界被钳位
 *   16#0003_013A【信息级】重试次数越界被钳位
 *   16#0003_02F0【故障级·组态使用类】未初始化、忙时重入或写入内容非法
 *   16#0003_02F1【故障级·组态类】超时重试耗尽
 *   16#0003_02F2【故障级·工艺类】读写头报错重试耗尽
 *   16#0003_02F3【故障级·工艺类】写后回读校验不符或非法状态兜底
 * 验收向量 (Acceptance) :
 *   V1 读链：就绪后调 ReadTag → 请求下发、忙态 → 硬件完成一拍并给出标签号
 *      → 读成功脉冲单拍、标签快照更新、读计数加 1
 *   V2 防重复读：抑制窗内再读到同一标签 → 不产生成功脉冲，置 0138；
 *      超过窗口后同一标签可再次成功
 *   V3 无标签：完成但标签号为空 → bNoTag 为 TRUE、bError 为 FALSE、
 *      重试计数不增不减
 *   V4 超时重试链：不给完成信号，重试上限 2 → 共 3 次下发后锁 02F1
 *   V5 写校验：写入后回读内容不一致 → 锁 02F3，写成功脉冲不产生
 *   V6 忙时重入：执行中再调读方法 → 返回 FALSE 并置 02F0
 *   V7 保持语义：读成功后停 10 拍，标签快照仍有效且内容不变
 * 红线自检 (Redline)    : R1 零全局变量表与外部变量引用 ｜ R2 零物理地址直写
 *                         R3 纯 IEC 61131-3 ｜ R4 字符串判等有注释说明（非浮点）、
 *                         计时器有界、无除法 ｜ R5 全变量中英双语同行注释
 *                         R6 ENUM 加 CASE 加 ELSE 兜底 ｜ R7 TON 与 R_TRIG 全部
 *                         在 CASE 之外无条件刷新
 * 修订历史 (Revision)   :
 *   2026-11-15  v1.0.0  首版入库（Round 10 · T2-6 Rockwell AOI 开组）
 *   2026-11-15  v1.0.1  R10 终审修复两处：
 *                       R-FIX-1【中等】uHwErrorCode 入参声明后从未使用，规格
 *                       要求的「读写头原始错误码透传进诊断」实际缺失；改为在
 *                       硬件报错拍写入诊断，并让段 9 的码刷新仅在块级码非零时
 *                       发生，避免每拍把透传值清成 0；
 *                       R-FIX-2【注释级】由此同步了诊断字段的真实刷新规则。
 * 规格偏离登记 (Deviations):
 *   D1 接口方法 Init 的 VAR_IN_OUT 形参名 stCfg 与本块 VAR_IN_OUT 引脚 stCfg
 *      同名（规格书两处都叫 stCfg），方法体内形参遮蔽同名引脚且方法体不引用
 *      形参，实际组态以块级引脚为准。改形参名会破坏 I_DL_RfidReader 契约，
 *      故按「契约优先」保留，现场联调务必把同一份组态实例同时接到引脚与
 *      Init 调用上（同一实例时二者天然一致）。
 *   D2 bHwReq / bHwWr 由规格书的内部 VAR 提为 VAR_OUTPUT：它们是送协议层或
 *      IO 层的指令电平，必须可被外部观测与接线，属向后兼容的可见性扩展。
 *============================================================================*)

(*------------------------------------------------------------------------------
 * 枚举: E_DL_RfidFsm（归属功能块 FB_DL_RfidTagHandler，与其同文件发布）
 * 内部五态，经属性 State 按写死的映射表折算为接口的五态
 *-----------------------------------------------------------------------------*)
TYPE E_DL_RfidFsm :
(
    eIdle   := 0,     // 待机：可受理请求 / Idle, accepts requests
    eWaitHw := 10,    // 已下发，等完成、报错或超时 / Command issued, waiting for done, error or timeout
    eVerify := 20,    // 写后回读校验 / Read-back verification after a write
    eRetry  := 30,    // 重试退避，单拍停留后重新下发 / Retry back-off, one cycle dwell then re-issue
    eFault  := 99     // 故障锁定，仅复位可退 / Fault latched, only reset leaves
);
END_TYPE

(*------------------------------------------------------------------------------
 * 枚举: E_DL_RfidReq（挂起请求类型，单发登记，消费即清）
 *-----------------------------------------------------------------------------*)
TYPE E_DL_RfidReq :
(
    eNone  := 0,      // 无挂起请求 / No pending request
    eRead  := 1,      // 挂起读标签请求 / Pending read request
    eWrite := 2       // 挂起写数据区请求 / Pending write request
);
END_TYPE

FUNCTION_BLOCK FB_DL_RfidTagHandler IMPLEMENTS I_DL_RfidReader
VAR_INPUT
    bEnable      : BOOL := TRUE;      // 使能，FALSE 转离线并拒绝全部方法 [-] / Enable, FALSE goes offline and rejects every method
    bHwReady     : BOOL;              // 读写头就绪反馈，由协议层或 IO 层注入 [-] / Reader ready feedback injected by the transport layer
    bHwDone      : BOOL;              // 本次指令执行完成，单拍或电平，内部取上升沿 [-] / Command done feedback, edge detected internally
    bHwError     : BOOL;              // 读写头报错反馈 [-] / Reader error feedback
    sHwTagId     : STRING(64);        // 读回的标签唯一号，空串表示视野内无标签 [ASCII] / Tag identifier read back, empty means no tag
    sHwData      : STRING(64);        // 读回的数据区内容 [ASCII 或十六进制] / Data area content read back
    uHwErrorCode : UDINT;             // 读写头原始错误码，透传进诊断不改语义 [代码] / Raw reader error code forwarded into diagnostics
    tCmdTimeout  : TIME := T#500MS;   // 单指令超时，域 50 毫秒到 5 秒 [毫秒] / Per-command timeout, 50 ms to 5 s
    nMaxRetry    : INT := 2;          // 重试次数，域 0 到 5 [次] / Retry count, 0 to 5
    bDupFilterEn : BOOL := TRUE;      // 同标签重复读抑制使能 [-] / Duplicate-read suppression enable
    tDupWindow   : TIME := T#2S;      // 重复读抑制窗，域 100 毫秒到 60 秒 [毫秒] / Duplicate suppression window
END_VAR
VAR_OUTPUT
    bReadDoneOk  : BOOL;              // 读成功，单拍脉冲 [-] / Read succeeded, single-cycle pulse
    bWriteDoneOk : BOOL;              // 写成功，单拍脉冲 [-] / Write succeeded, single-cycle pulse
    bNoTag       : BOOL;              // 视野内无标签，保持型业务态 [-] / No tag in field, holding business state
    bBusy        : BOOL;              // 指令执行中 [-] / Command in progress
    bError       : BOOL;              // 故障锁存，组态类与工艺类同置，码区分 [-] / Fault latch, both classes set it, the code tells them apart
    uErrorId     : UDINT;             // 事件码，0 = 无事件 / Event code, 0 = no event
    nRetryCnt    : INT;               // 本次指令已重试次数 [次] / Retries already spent on the current command
    bHwReq       : BOOL;              // 硬件请求电平，送协议层或 IO 层 [-] / Hardware request level towards the transport layer
    bHwWr        : BOOL;              // 硬件读写方向，FALSE 为读，TRUE 为写 [-] / Direction towards the hardware, FALSE reads, TRUE writes
END_VAR
VAR_IN_OUT
    stCfg        : ST_DL_RfidCfg;     // 组态，调用方持有，本块只读使用 [结构] / Configuration owned by the caller, read-only here
END_VAR
VAR
    fbTrigDone   : R_TRIG;            // 硬件完成沿检测，CASE 之外无条件刷新 [-] / Rising edge detector for the hardware done signal
    fbTmo        : TON;               // 单指令超时计时，CASE 之外无条件刷新 [-] / Command timeout timer refreshed outside the CASE
    fbDupTmo     : TON;               // 重复读抑制窗计时，栅极复位 [-] / Duplicate suppression window timer with gate reset
    fbAge        : TON;               // 通信年龄计时，成功时栅极复位 [-] / Communication age timer reset on success
    bInit        : BOOL := FALSE;     // 首扫标志，初值 FALSE，判据 NOT bInit（R19 范式）[-] / First-scan flag
    bInitDone    : BOOL;              // 已收到 Init 请求且组态已装载 [-] / TRUE after a successful Init request
    eState       : E_DL_RfidFsm := E_DL_RfidFsm.eIdle;  // 内部主状态机 / Internal main state machine
    eReq         : E_DL_RfidReq := E_DL_RfidReq.eNone;  // 挂起请求类型 / Pending request type
    bReqInit     : BOOL;              // Init 方法登记的单发请求 [-] / Single-shot request registered by the Init method
    bReqReset    : BOOL;              // Reset 方法登记的单发请求 [-] / Single-shot request registered by the Reset method
    bTmoIn       : BOOL;              // 超时定时器输入条件，先算后调以免条件调用实例 [-] / Timer input condition computed before the unconditional call
    sLastTagId   : STRING(64);        // 上次成功读取的标签号，重复抑制比对源 [ASCII] / Last accepted tag identifier, the comparison source
    sWrBuffer    : STRING(64);        // 待写内容副本，防止调用方中途改动 [ASCII] / Latched write payload, immune to caller changes
    stTag        : ST_DL_RfidTag;     // 当前标签快照，属性出口 [-] / Current tag snapshot served by the Tag property
    stDiag       : ST_DL_RfidDiag;    // 诊断结构，属性出口 [-] / Diagnostic structure served by the Diag property
    bDupGate     : BOOL := TRUE;      // 重复窗计时栅极，接受标签后拉低一拍 [-] / Gate of the duplicate timer, pulled low for one cycle on accept
    bDupRearm    : BOOL;              // 重复窗栅极再武装标志 [-] / Re-arm flag of the duplicate timer gate
    bAgeGate     : BOOL := TRUE;      // 通信年龄计时栅极，成功后拉低一拍 [-] / Gate of the age timer, pulled low for one cycle on success
    bAgeRearm    : BOOL;              // 通信年龄栅极再武装标志 [-] / Re-arm flag of the age timer gate
    tTmoUse      : TIME := T#500MS;   // 生效超时（已仲裁与钳位）[毫秒] / Effective timeout after arbitration and clamping
    tDupUse      : TIME := T#2S;      // 生效抑制窗（已仲裁与钳位）[毫秒] / Effective suppression window after arbitration and clamping
    nRetryUse    : INT := 2;          // 生效重试次数（已仲裁与钳位）[次] / Effective retry count after arbitration and clamping
    bDupUse      : BOOL := TRUE;      // 生效重复抑制使能 [-] / Effective duplicate suppression enable
    bLastTimeout : BOOL;              // 上次失败是否为超时，用于区分耗尽码 [-] / TRUE when the last failure was a timeout
END_VAR
VAR CONSTANT
    DL_RFID_TMO_MIN   : TIME := T#50MS;    // 超时下限 [毫秒] / Timeout lower bound
    DL_RFID_TMO_MAX   : TIME := T#5S;      // 超时上限 [毫秒] / Timeout upper bound
    DL_RFID_DUP_MIN   : TIME := T#100MS;   // 抑制窗下限 [毫秒] / Suppression window lower bound
    DL_RFID_DUP_MAX   : TIME := T#60S;     // 抑制窗上限 [毫秒] / Suppression window upper bound
    DL_RFID_RETRY_MAX : INT  := 5;         // 重试上限 [次] / Retry upper bound
    DL_RFID_RETRY_MIN : INT  := 0;         // 重试下限，0 表示不重试 [次] / Retry lower bound, zero means no retry
    DL_STR_MAX        : INT  := 64;        // 字符串域长度上限，与 STRING(64) 一致 [字符] / String capacity, kept in sync with STRING(64)
    DL_RFID_AGE_MAX   : TIME := T#24H;     // 通信年龄计时上限，超时后停在终点值 [毫秒] / Age timer span ceiling
END_VAR

METHOD Init : BOOL
VAR_IN_OUT
    stCfg : ST_DL_RfidCfg;    // 组态结构，调用方持有，本方法只登记不阻塞 [结构] / Configuration injected by the caller
END_VAR
Init := FALSE;
IF NOT bEnable THEN
    stDiag.uLastErrorId := 16#0003_02F0;    // 失能状态下拒绝初始化
    RETURN;
END_IF
bReqInit := TRUE;                            // 只登记，装载在主体段 6 执行
Init     := TRUE;

(*------------------------------------------------------------------------------
 * 方法实现：ReadTag（单发登记，忙时拒绝且不排队）
 *      Method ReadTag: single-shot registration, rejected while busy, never queued
 *-----------------------------------------------------------------------------*)
    END_METHOD

METHOD ReadTag : BOOL
VAR_INPUT
END_VAR
ReadTag := FALSE;
IF NOT bEnable THEN
    stDiag.uLastErrorId := 16#0003_02F0;
    RETURN;
END_IF
IF NOT bInitDone THEN
    stDiag.uLastErrorId := 16#0003_02F0;    // 未初始化：拒绝
    RETURN;
END_IF
IF eState <> E_DL_RfidFsm.eIdle THEN
    stDiag.uLastErrorId := 16#0003_02F0;    // 忙时重入：拒绝，不排队
    RETURN;
END_IF
IF eReq <> E_DL_RfidReq.eNone THEN
    stDiag.uLastErrorId := 16#0003_02F0;    // 已有挂起请求：拒绝，避免覆盖
    RETURN;
END_IF
eReq    := E_DL_RfidReq.eRead;
ReadTag := TRUE;

(*------------------------------------------------------------------------------
 * 方法实现：WriteTag（单发登记 + 内容副本锁存）
 *      Method WriteTag: single-shot registration with a latched payload copy
 *      字符串长度越界：STRING(64) 已由编译器保证长度，故本分支退化为
 *      「空内容拒绝」，并在头注释与本段注释双重声明（R11 留档）
 *-----------------------------------------------------------------------------*)
    END_METHOD

METHOD WriteTag : BOOL
VAR_IN_OUT
    stTagIn : ST_DL_RfidTag;    // 待写内容，本方法立即拷贝到内部缓冲 [结构] / Payload latched into the internal buffer
END_VAR
WriteTag := FALSE;
IF NOT bEnable THEN
    stDiag.uLastErrorId := 16#0003_02F0;
    RETURN;
END_IF
IF NOT bInitDone THEN
    stDiag.uLastErrorId := 16#0003_02F0;
    RETURN;
END_IF
IF eState <> E_DL_RfidFsm.eIdle THEN
    stDiag.uLastErrorId := 16#0003_02F0;    // 忙时重入：拒绝
    RETURN;
END_IF
IF eReq <> E_DL_RfidReq.eNone THEN
    stDiag.uLastErrorId := 16#0003_02F0;
    RETURN;
END_IF
IF stTagIn.sData = '' THEN
    stDiag.uLastErrorId := 16#0003_02F0;    // 空内容等同于写入长度非法
    RETURN;
END_IF
sWrBuffer := stTagIn.sData;                  // 立即拷贝，防调用方中途改动
eReq      := E_DL_RfidReq.eWrite;
WriteTag  := TRUE;

(*------------------------------------------------------------------------------
 * 方法实现：Reset（故障态下唯一受理的方法）
 *      Method Reset: the only method accepted in the fault state
 *-----------------------------------------------------------------------------*)
    END_METHOD

METHOD Reset : BOOL
VAR_INPUT
END_VAR
Reset     := TRUE;
bReqReset := TRUE;

(*------------------------------------------------------------------------------
 * 属性实现（R22：接口成员一律只读 PROPERTY GET）
 *      Property implementations, read-only GET as required by the interface
 *-----------------------------------------------------------------------------*)
    END_METHOD

(*------------------------------------------------------------------------------
 * 段 1｜单拍输出预清零（R25 律①）：两个成功脉冲必须在主体最前部清零
 *      Single-cycle output pre-clear: both success pulses cleared at the very top
 *-----------------------------------------------------------------------------*)
bReadDoneOk  := FALSE;
bWriteDoneOk := FALSE;

(*------------------------------------------------------------------------------
 * 段 2｜完成沿检测（R7 红线）：实例在 CASE 之外无条件刷新
 *      Done edge detection, instance refreshed outside any branch
 *-----------------------------------------------------------------------------*)
fbTrigDone(CLK := bHwDone);

(*------------------------------------------------------------------------------
 * 段 3｜首扫初始化（R19 唯一合法范式）
 *      First-scan initialisation with the canonical R19 pattern
 *-----------------------------------------------------------------------------*)
IF NOT bInit THEN
    eState     := E_DL_RfidFsm.eIdle;
    eReq       := E_DL_RfidReq.eNone;
    nRetryCnt  := 0;
    bError     := FALSE;
    uErrorId   := 16#0000_0000;
    bNoTag     := FALSE;
    bInitDone  := FALSE;
    sLastTagId := '';
    sWrBuffer  := '';
    stTag.sTagId := '';
    stTag.sData  := '';
    stTag.uPage  := 0;
    stTag.nRssi  := 0;
    stTag.bValid := FALSE;
    stDiag.uLastErrorId := 0;
    stDiag.nCommRetry   := 0;
    stDiag.nReadTotal   := 0;
    stDiag.nWriteTotal  := 0;
    stDiag.bAntennaOk   := FALSE;
    stDiag.tLastComm    := T#0S;
    bInit      := TRUE;                  // 首扫只做一次
END_IF

(*------------------------------------------------------------------------------
 * 段 4｜组态仲裁与钳位（三源优先级写死：常量域 低于 引脚 低于 Init 组态）
 *      Configuration arbitration with a fixed three-level priority
 *      同一字段只沿一个方向回落，不出现隐式切换；越界一律钳位并置 0139 或 013A
 *-----------------------------------------------------------------------------*)
IF bInitDone AND (stCfg.tTimeout >= DL_RFID_TMO_MIN) AND (stCfg.tTimeout <= DL_RFID_TMO_MAX) THEN
    tTmoUse := stCfg.tTimeout;
ELSE
    tTmoUse := tCmdTimeout;
END_IF
IF tTmoUse < DL_RFID_TMO_MIN THEN
    tTmoUse  := DL_RFID_TMO_MIN;
    uErrorId := 16#0003_0139;
ELSIF tTmoUse > DL_RFID_TMO_MAX THEN
    tTmoUse  := DL_RFID_TMO_MAX;
    uErrorId := 16#0003_0139;
END_IF

IF bInitDone AND (stCfg.tDupWindow >= DL_RFID_DUP_MIN) AND (stCfg.tDupWindow <= DL_RFID_DUP_MAX) THEN
    tDupUse := stCfg.tDupWindow;
ELSE
    tDupUse := tDupWindow;
END_IF
IF tDupUse < DL_RFID_DUP_MIN THEN
    tDupUse  := DL_RFID_DUP_MIN;
    uErrorId := 16#0003_0139;
ELSIF tDupUse > DL_RFID_DUP_MAX THEN
    tDupUse  := DL_RFID_DUP_MAX;
    uErrorId := 16#0003_0139;
END_IF

IF bInitDone THEN
    nRetryUse := stCfg.nMaxRetry;
ELSE
    nRetryUse := nMaxRetry;
END_IF
IF nRetryUse < DL_RFID_RETRY_MIN THEN
    nRetryUse := DL_RFID_RETRY_MIN;
    uErrorId  := 16#0003_013A;
ELSIF nRetryUse > DL_RFID_RETRY_MAX THEN
    nRetryUse := DL_RFID_RETRY_MAX;
    uErrorId  := 16#0003_013A;
END_IF

IF bInitDone THEN
    bDupUse := stCfg.bDupFilterEn;
ELSE
    bDupUse := bDupFilterEn;
END_IF

(*------------------------------------------------------------------------------
 * 段 5｜计时器无条件周期刷新（红线第 7 条）：三个 TON 全部在 CASE 之外
 *      All three timers refreshed outside the CASE, mandatory by the red line
 *      单指令超时：IN 条件先算进 bTmoIn，再无条件调用实例，禁止把调用写进 IF
 *-----------------------------------------------------------------------------*)
IF eState = E_DL_RfidFsm.eWaitHw THEN
    bTmoIn := TRUE;
ELSE
    bTmoIn := FALSE;
END_IF
fbTmo(IN := bTmoIn, PT := tTmoUse);

(* 重复抑制窗：栅极拉低一整拍才能复位 TON，再武装标志在调用之后置回高电平 *)
fbDupTmo(IN := bDupGate AND bDupUse, PT := tDupUse);
IF bDupRearm THEN
    bDupRearm := FALSE;
    bDupGate  := TRUE;
END_IF

(* 通信年龄：成功一次即复位并重新计时，用于诊断「多久没读到东西」 *)
fbAge(IN := bAgeGate, PT := DL_RFID_AGE_MAX);
IF bAgeRearm THEN
    bAgeRearm := FALSE;
    bAgeGate  := TRUE;
END_IF

(*------------------------------------------------------------------------------
 * 段 6｜单发请求消费（Init 与 Reset）：置位 到 消费 到 复位，三律齐全
 *      Consume the Init and Reset single-shot requests, place, consume, clear
 *-----------------------------------------------------------------------------*)
IF bReqInit THEN
    bReqInit := FALSE;                       // 先复位标志，避免跨拍泄漏
    IF bEnable THEN
        bInitDone           := TRUE;
        stDiag.bAntennaOk   := TRUE;         // 天线由组态确认；实际自检由硬件层给
        stDiag.uLastErrorId := 0;
        uErrorId            := 16#0000_0000;
    END_IF
END_IF

IF bReqReset THEN
    bReqReset := FALSE;                      // 先复位标志
    bError    := FALSE;
    uErrorId  := 16#0000_0000;
    nRetryCnt := 0;
    bNoTag    := FALSE;
    bHwReq    := FALSE;
    eReq      := E_DL_RfidReq.eNone;
    eState    := E_DL_RfidFsm.eIdle;
END_IF

(*------------------------------------------------------------------------------
 * 段 7｜失能拦截（每拍最先判）：清请求与硬件请求，故障锁存保留
 *      Disable interception: clear requests and the hardware request, keep the latch
 *-----------------------------------------------------------------------------*)
IF NOT bEnable THEN
    bHwReq := FALSE;
    bBusy  := FALSE;
    eReq   := E_DL_RfidReq.eNone;
    IF eState <> E_DL_RfidFsm.eFault THEN
        eState := E_DL_RfidFsm.eIdle;
    END_IF
END_IF

(*------------------------------------------------------------------------------
 * 段 8｜主状态机（ENUM 加 CASE，含 ELSE 兜底）
 *      Main state machine with an ELSE fallback branch
 *-----------------------------------------------------------------------------*)
CASE eState OF
    E_DL_RfidFsm.eIdle:
        bHwReq := FALSE;
        IF bEnable AND bHwReady AND bInitDone AND (eReq <> E_DL_RfidReq.eNone) THEN
            IF eReq = E_DL_RfidReq.eWrite THEN
                bHwWr := TRUE;               // 写方向
            ELSE
                bHwWr := FALSE;              // 读方向
            END_IF
            bHwReq       := TRUE;            // 下发请求（电平，硬件层取上升沿）
            nRetryCnt    := 0;               // 新指令重试计数清零
            bNoTag       := FALSE;           // 新指令开始清业务态
            bLastTimeout := FALSE;
            eState       := E_DL_RfidFsm.eWaitHw;
        END_IF

    E_DL_RfidFsm.eWaitHw:
        bHwReq := TRUE;                      // 保持请求电平直到有结论
        IF fbTrigDone.Q THEN
            IF bHwError THEN
                (* 读写头报错：走重试链，耗尽按工艺类 02F2 报
                   硬件原始码在此处原样透传进诊断（不改语义），现场据此查手册；
                   耗尽后 uLastErrorId 会记块级码 02F2，原始码仍可经 uHwErrorCode
                   引脚读取，两级信息都不丢 *)
                stDiag.uLastErrorId := uHwErrorCode;
                bLastTimeout := FALSE;
                bHwReq       := FALSE;
                eState       := E_DL_RfidFsm.eRetry;
            ELSIF sHwTagId = '' THEN
                (* 无标签：业务态，不计重试、不置故障 *)
                bNoTag := TRUE;
                eReq   := E_DL_RfidReq.eNone;
                bHwReq := FALSE;
                eState := E_DL_RfidFsm.eIdle;
            ELSIF eReq = E_DL_RfidReq.eRead THEN
                IF bDupUse AND (sHwTagId = sLastTagId) AND (NOT fbDupTmo.Q) THEN
                    (* 抑制窗内同一标签：丢弃结果，只记信息级码 *)
                    uErrorId := 16#0003_0138;
                    eReq     := E_DL_RfidReq.eNone;
                    bHwReq   := FALSE;
                    eState   := E_DL_RfidFsm.eIdle;
                ELSE
                    (* 正常读取：锁存快照并置单拍成功脉冲 *)
                    stTag.sTagId := sHwTagId;
                    stTag.sData  := sHwData;
                    stTag.uPage  := 0;
                    stTag.nRssi  := 0;
                    stTag.bValid := TRUE;
                    sLastTagId   := sHwTagId;
                    stDiag.nReadTotal := stDiag.nReadTotal + 1;
                    bReadDoneOk  := TRUE;
                    bDupGate     := FALSE;   // 抑制窗从零重新计时
                    bDupRearm    := TRUE;
                    bAgeGate     := FALSE;   // 通信年龄从零重新计时
                    bAgeRearm    := TRUE;
                    eReq         := E_DL_RfidReq.eNone;
                    bHwReq       := FALSE;
                    eState       := E_DL_RfidFsm.eIdle;
                END_IF
            ELSE
                (* 写请求完成：转回读校验态，不在本态直接报成功 *)
                bHwWr  := TRUE;
                eState := E_DL_RfidFsm.eVerify;
            END_IF
        ELSIF fbTmo.Q THEN
            (* 超时：走重试链，耗尽按组态类 02F1 报 *)
            bLastTimeout := TRUE;
            bHwReq       := FALSE;
            eState       := E_DL_RfidFsm.eRetry;
        END_IF

    E_DL_RfidFsm.eVerify:
        (* 写后回读校验：字符串判等合法（字符串不是浮点数，不存在容差问题） *)
        bHwReq := FALSE;
        IF sHwData = sWrBuffer THEN
            stTag.sData  := sWrBuffer;
            stTag.bValid := TRUE;
            stDiag.nWriteTotal := stDiag.nWriteTotal + 1;
            bWriteDoneOk := TRUE;
            bAgeGate     := FALSE;
            bAgeRearm    := TRUE;
            eReq         := E_DL_RfidReq.eNone;
            eState       := E_DL_RfidFsm.eIdle;
        ELSE
            uErrorId := 16#0003_02F3;        // 工艺类：回读不符
            bError   := TRUE;
            eReq     := E_DL_RfidReq.eNone;
            eState   := E_DL_RfidFsm.eFault;
        END_IF

    E_DL_RfidFsm.eRetry:
        (* 退避单拍：请求电平拉低一拍，重新下发时自然形成新的上升沿 *)
        bHwReq    := FALSE;
        nRetryCnt := nRetryCnt + 1;
        IF nRetryCnt > nRetryUse THEN
            IF bLastTimeout THEN
                uErrorId := 16#0003_02F1;    // 组态类：超时重试耗尽
            ELSE
                uErrorId := 16#0003_02F2;    // 工艺类：读写头报错重试耗尽
            END_IF
            bError := TRUE;
            eReq   := E_DL_RfidReq.eNone;
            eState := E_DL_RfidFsm.eFault;
        ELSE
            eState := E_DL_RfidFsm.eWaitHw;  // 重新下发，请求域沿用锁存值
        END_IF

    E_DL_RfidFsm.eFault:
        (* 故障锁定：请求电平清零，退出只能靠 Reset 方法（段 6 已消费） *)
        bHwReq := FALSE;

    ELSE
        (* 非法枚举值兜底 *)
        eState   := E_DL_RfidFsm.eFault;
        uErrorId := 16#0003_02F3;
        bError   := TRUE;
        bHwReq   := FALSE;
END_CASE

(*------------------------------------------------------------------------------
 * 段 9｜派生输出与诊断每拍重写（R27）
 *      Derived outputs and diagnostics rewritten every cycle
 *-----------------------------------------------------------------------------*)
IF eState = E_DL_RfidFsm.eFault THEN
    bError := TRUE;              // 故障锁存：进入故障态即置位，退出只能靠 Reset
END_IF

IF (eState = E_DL_RfidFsm.eWaitHw) OR (eState = E_DL_RfidFsm.eVerify) OR (eState = E_DL_RfidFsm.eRetry) THEN
    bBusy := TRUE;
ELSE
    bBusy := FALSE;
END_IF

stDiag.nCommRetry   := nRetryCnt;
IF uErrorId <> 16#0000_0000 THEN
    stDiag.uLastErrorId := uErrorId;   // 仅在块级码非零时刷新，避免把透传的硬件原始码清掉
END_IF
stDiag.tLastComm    := fbAge.ET;

(*------------------------------------------------------------------------------
 * 方法实现：Init（单发登记 + 组态注入）
 *      Method Init: single-shot registration with configuration injection
 *-----------------------------------------------------------------------------*)

PROPERTY State : E_DL_RfidState
(* 映射写死，禁止就近映射：无标签业务态优先级最高，其次故障，其次离线，最后忙态 *)
IF bNoTag THEN
    State := E_DL_RfidState.eNoTag;
ELSIF eState = E_DL_RfidFsm.eFault THEN
    State := E_DL_RfidState.eError;
ELSIF (NOT bEnable) OR (NOT bInitDone) OR (NOT bHwReady) THEN
    State := E_DL_RfidState.eOffline;
ELSIF eState = E_DL_RfidFsm.eIdle THEN
    State := E_DL_RfidState.eReady;
ELSE
    State := E_DL_RfidState.eBusy;
END_IF

PROPERTY Tag : ST_DL_RfidTag
Tag := stTag;                    // 保持型快照（R27），直到下次成功读取覆盖

PROPERTY Diag : ST_DL_RfidDiag
Diag := stDiag;                  // 诊断整体回读，等价于 AOI 的 InOut 段封装
END_FUNCTION_BLOCK

(* ---- FB_DL_SafetyLightCurtain.st ---- *)
(*==============================================================================
 * 组件名称 (Component)  : FB_DL_SafetyLightCurtain
 * 所属子库 (Sublibrary) : DL_Device
 * 当前版本 (Version)    : 1.0.1
 * 兼容性   (Platform)   : CODESYS 3.5 / TwinCAT 3 / 汇川 InoProShop / Machine Expert
 *                         仅依赖 Standard.library（TON / R_TRIG），零厂商方言
 * 分类     (Category)   : 设备功能块（Function Block，实现 I_DL_LightCurtain）
 * 功能简述 (Function)   : 光幕 OSSD 监控 + 2/4 传感器序列屏蔽状态机 + 屏蔽
 *                         总时长超时 + 滞留清除 override + 屏蔽灯输出（屏蔽
 *                         常亮/override 闪烁）+ 故障复位联锁（SICK mut_p /
 *                         西门子 Sequential Muting 公开语义 clean-room）。
 * 定位声明 (Positioning): 公约 0.13——本块为标准 PLC 逻辑编排与诊断镜像层，
 *                         不构成 ISO 13849 / IEC 62061 认证安全功能，安全回
 *                         路由认证安全控制器/安全 PLC 承载；光幕本体 OSSD
 *                         的安全判断在认证安全光幕内部完成，本块仅做诊断镜
 *                         像与屏蔽编排。
 * 接口实现 (Implements) : I_DL_LightCurtain。接口属性同名成员（eState/bClear/
 *                         bMutingActive/bOverrideActive/bSafeStop/bFault/
 *                         uErrorId）按 R22 以只读 PROPERTY GET 承载（内部镜
 *                         像同源），非接口成员 bMutingLamp 保留 VAR_OUTPUT；
 *                         方法 CmdOverride/CmdAck/CmdReset 在本文件尾部落地。
 * 公约遵循 (Convention) : 0.1/R23 事件/电平混合编排（电平条件级联驱动，无连
 *                         续量同步语义），免首扫，无 bInit。
 *                         0.2/R21 bFault 显式排除信息级码；0.5/R7 全部实例主
 *                         体最前部无条件刷新；0.7/R15 故障级锁存仅复位路径
 *                         清码。
 *                         0.8 故障码段位 16#0003_xxxx（经 DL_Device
 *                         VERSION.md 码表核对：规格建议 0003_0270/0271/0272
 *                         已被 FB_DL_ThreePointValve 占用、0003_0106 已被
 *                         FB_DL_VfdGeneric 占用，依公约冲突顺延）：
 *                         【故障级】0003_02A0 屏蔽传感器序列错误、0003_02A1
 *                         屏蔽超时、0003_02A2 OSSD 双通道不一致；
 *                         【信息级】0003_0122 override 准入拒绝（无遮挡）、
 *                         0003_0118 override 硬帽到期退出。
 * 红线自检 (Redline)    : R1 零全局变量表/外部变量引用 ✓｜R2 零物理 IO 地址 ✓
 *                         R3 纯 IEC 61131-3 ✓｜R4 参数钳位/超窗防御 ✓
 *                         R5 全变量中英双语同行注释 ✓｜R6 状态映像 IF 派生
 *                         链含 ELSE 兜底（无显式 CASE 主状态机，见偏离①）✓
 *                         R7 五实例（R_TRIG×1/TON×4）主体最前部无条件刷新 ✓
 *                         R8 全常量化 ✓
 * 设计要点 (Key notes)  : ① 序列屏蔽：2 传感器 M1→M2 进入、M1→M2 清离退出；
 *                           4 传感器正向 M1→M2 进入、M3→M4 离开、全清退出，
 *                           反向全程镜像；序列错乱 → 立即退出屏蔽 + 故障 +
 *                           bSafeStop 按光幕实际状态输出；
 *                         ② override 准入硬约束：bOverrideKey（或方法请求）
 *                           AND 屏蔽传感器至少一真才进入，无遮挡拒绝置信级；
 *                         ③ 屏蔽灯闪烁用主周期 TON 振荡器自实现（方波生成
 *                           不用 TON 单实例直出，用 IN:=NOT Q 重触发振荡法；
 *                           R14 断输入一拍规则不涉及方波生成，注释说明）；
 *                         ④ OSSD 双通道不一致超 tDiscrepancy → 故障锁存；
 *                         ⑤ bSafeStop 出口断言：屏蔽/override 态恒 FALSE
 *                           （光幕正常），永不因屏蔽置假。
 * 偏离留档 (Deviation)  : 依 R11 头注释留档，共 2 条：
 *                         ① 码位与兜底态：规格建议 0003_0270/0271/0272/0273
 *                           与既有 FB_DL_ThreePointValve 冲突，顺延为
 *                           0003_02A0/02A1/02A2；因本块状态为条件派生映像
 *                           （无独立 CASE 主状态机），「非法状态兜底」码不
 *                           适用而取消，派生链含 ELSE 兜底保证域外输入归安
 *                           全侧（核对结果优先于建议值）。
 *                         ② 反向序列：2 传感器模式以「首遮挡传感器」判定方
 *                           向（M1 先遮挡=正向）；4 传感器模式同理（M4 先
 *                           遮挡=反向），方向一经判定锁定至本序列结束。
 * 开源溯源 (Origin)     : 来源标签 tcopen-component / light-curtain-muting
 *                         （RAW_NOTES_R7 S-5：SICK mut_p 与西门子 Sequential
 *                         Muting 公开手册语义——2/4 传感器序列、容差窗、
 *                         override 硬帽、屏蔽灯，公开资料，仅借鉴语义域；
 *                         状态步进实现、码位与引脚契约 100% 本库独立设计，
 *                         clean-room 未复制源码）。
 * 验收向量 (Acceptance) :
 *   V1 无屏蔽遮挡停机链：光幕遮挡且未屏蔽 → bSafeStop=TRUE、eState=eBlocked；
 *   V2 2 传感器合法序列：M1→M2 遮挡（屏蔽灯常亮，bSafeStop=FALSE）→ M1 清
 *      → M2 清（序列完成回 eClear）；
 *   V3 序列错乱停机：M2 先遮挡后 M1 清（E2 清而 E1 仍遮挡）→ 故障 0003_02A0
 *      + bSafeStop 按实际 OSSD 输出；
 *   V4 屏蔽超时：序列驻留超 tMutingTimeout → 故障 0003_02A1；
 *   V5 override 准入/拒绝/硬帽：钥匙开关无遮挡 → 拒绝置信级 0003_0122；有遮
 *      挡 → eOverride 灯闪；超 tOverrideMax → 退出 + 0003_0118；
 *   V6 OSSD 不一致：双通道异电平超 tDiscrepancy → 故障 0003_02A2；
 *   V7 复位联锁：故障后仅 bReset 沿且故障源消失才解除锁存。
 * 修订历史 (Revision)   :
 *   2026-11-15  v1.0.0  首版入库（Round 07 · DL_Device 光幕族实现件）
 *   2026-11-15  v1.0.1  终审修复 2 处：① 反向序列判向条件与偏离②矛盾——
 *                       2 传感器模式判向 ELSIF 与正向 IF 恒等（死代码）、4
 *                       传感器模式误查 M3（应为 M4=_bX2），按「M2/M4 先遮挡=
 *                       反向」修正；② 2 传感器 E2 步双清离无分支 → 步号滞留、
 *                       依赖屏蔽超时误报故障，补双清离回 IDLE（中断恢复）
 *============================================================================*)
FUNCTION_BLOCK FB_DL_SafetyLightCurtain IMPLEMENTS I_DL_LightCurtain
VAR_INPUT
    bOssd1          : BOOL;             // 光幕 OSSD 通道 1（OSSD channel 1），TRUE=通光 / OSSD channel 1, TRUE = clear
    bOssd2          : BOOL;             // 光幕 OSSD 通道 2（OSSD channel 2），TRUE=通光 / OSSD channel 2, TRUE = clear
    bMutSens1       : BOOL;             // 屏蔽传感器 1（Muting sensor 1），TRUE=被遮挡；2 传感器模式使用 / Muting sensor 1, TRUE = blocked, 2-sensor mode
    bMutSens2       : BOOL;             // 屏蔽传感器 2（Muting sensor 2），TRUE=被遮挡；2 传感器模式使用 / Muting sensor 2, TRUE = blocked, 2-sensor mode
    bMutSens3       : BOOL;             // 屏蔽传感器 3（Muting sensor 3），TRUE=被遮挡；4 传感器模式使用 / Muting sensor 3, TRUE = blocked, 4-sensor mode
    bMutSens4       : BOOL;             // 屏蔽传感器 4（Muting sensor 4），TRUE=被遮挡；4 传感器模式使用 / Muting sensor 4, TRUE = blocked, 4-sensor mode
    bFourSensorMode : BOOL;             // 四传感器模式选择（Four-sensor mode），TRUE=序列式 4 传感器；FALSE=2 传感器 / TRUE = 4-sensor sequential, FALSE = 2-sensor
    bEnableMuting   : BOOL;             // 屏蔽功能总使能（Muting enable），FALSE=任何屏蔽条件都不生效（纯防护模式）/ FALSE disables all muting, pure guard mode
    bOverrideKey    : BOOL;             // 滞留清除钥匙开关（Override key，双通道语义由接线层保证），电平保持式 / Override key, level-held
    bReset          : BOOL;             // 复位按钮（Reset），上升沿复位故障与重启联锁 / Reset edge clears fault and restart interlock
    tMutingTimeout  : TIME := T#30S;    // 屏蔽总时长上限（Muting timeout），域 1S~600S 越界钳位；首末传感器间隔超限即故障 / Muting total-time cap, clamped 1S..600S
    tDiscrepancy    : TIME := T#3S;     // 传感器容差窗（Sensor discrepancy time），域 100MS~10S 越界钳位 / Discrepancy window, clamped 100MS..10S
    tOverrideMax    : TIME := T#30S;    // 滞留清除硬帽（Override max time），域 1S~60S 越界钳位 / Override hard cap, clamped 1S..60S
END_VAR
VAR_OUTPUT
    bMutingLamp : BOOL;                 // 屏蔽灯输出（Muting lamp）：屏蔽常亮、override 闪烁 / Muting lamp: steady in muting, blinking in override
END_VAR
VAR
    _eState       : E_DL_CurtainState;  // 派生状态映像（Derived state image），属性只读 / Derived state, read-only via property
    _bFaultLatch  : BOOL;               // 故障锁存标志（Fault latch flag），仅复位路径清除 / Fault latch, cleared only via reset path
    _uErrorIdInt  : UDINT;              // 内部故障级码寄存（Internal fault-level register）/ Internal fault-level register
    _uInfoCode    : UDINT;              // 本拍信息级码（Info code this cycle），瞬时型每拍重算 / Transient info code, recomputed each scan
    _nMutStep     : USINT;              // 屏蔽序列步号（Muting sequence step），0=空闲 / Muting step, 0 = idle
    _bMutRev      : BOOL;               // 反向序列方向标志（Reverse sequence direction），首遮挡传感器判定 / Reverse direction by first-blocked sensor
    _bE1          : BOOL;               // 映射后进入侧传感器 1（Mapped entry sensor 1）/ Mapped entry sensor 1
    _bE2          : BOOL;               // 映射后进入侧传感器 2（Mapped entry sensor 2）/ Mapped entry sensor 2
    _bX1          : BOOL;               // 映射后离开侧传感器 1（Mapped exit sensor 1）/ Mapped exit sensor 1
    _bX2          : BOOL;               // 映射后离开侧传感器 2（Mapped exit sensor 2）/ Mapped exit sensor 2
    _bMutingAct   : BOOL;               // 屏蔽进行中派生（Muting-active derived flag）/ Muting-active derived flag
    _bOverrideAct : BOOL;               // 滞留清除进行中（Override active flag）/ Override active flag
    _bPendOverride: BOOL;               // 方法 override 请求（Method override request）/ Method override request
    _bPendAck     : BOOL;               // 方法确认请求（Method ack request）/ Method ack request
    _bPendReset   : BOOL;               // 方法复位请求（Method reset request）/ Method reset request
    _bAnyMutBlocked: BOOL;              // 屏蔽传感器任一遮挡（Any muting sensor blocked）/ Any muting sensor blocked
    _tMutToEff    : TIME := T#30S;      // 钳位后屏蔽超时（Clamped muting timeout）/ Clamped muting timeout
    _tDiscEff     : TIME := T#3S;       // 钳位后容差窗（Clamped discrepancy window）/ Clamped discrepancy window
    _tOvrMaxEff   : TIME := T#30S;      // 钳位后 override 硬帽（Clamped override cap）/ Clamped override cap
    _fbTrigReset  : R_TRIG;             // 复位沿（Reset edge）/ Reset edge detector
    _fbTonDisc    : TON;                // OSSD 双通道容差窗（OSSD discrepancy window）/ OSSD discrepancy window
    _fbTonMutTo   : TON;                // 屏蔽总时长超时（Muting total-time timeout）/ Muting total-time timeout
    _fbTonOvrMax  : TON;                // override 硬帽计时（Override hard-cap timer）/ Override hard-cap timer
    _fbTonBlink   : TON;                // 屏蔽灯闪烁振荡器（Lamp blink oscillator），IN:=NOT Q 重触发 / Lamp blink oscillator, retriggered by NOT Q
END_VAR
VAR CONSTANT
    DL_BLINK_HALF : TIME := T#250MS;    // 屏蔽灯闪烁半周期（Lamp blink half period）/ Lamp blink half period
    DL_MUTTO_MIN  : TIME := T#1S;       // 屏蔽超时下限（Muting timeout lower clamp）/ Muting timeout lower clamp
    DL_MUTTO_MAX  : TIME := T#600S;     // 屏蔽超时上限（Muting timeout upper clamp）/ Muting timeout upper clamp
    DL_DISC_MIN   : TIME := T#100MS;    // 容差窗下限（Discrepancy lower clamp）/ Discrepancy lower clamp
    DL_DISC_MAX   : TIME := T#10S;      // 容差窗上限（Discrepancy upper clamp）/ Discrepancy upper clamp
    DL_OVR_MIN    : TIME := T#1S;       // override 硬帽下限（Override cap lower clamp）/ Override cap lower clamp
    DL_OVR_MAX    : TIME := T#60S;      // override 硬帽上限（Override cap upper clamp）/ Override cap upper clamp
    MUT_STEP_IDLE  : USINT := 0;        // 序列步：空闲（Step: idle）/ Step: idle
    MUT_STEP_E1    : USINT := 1;        // 序列步：首进入传感器已遮挡（Step: first entry sensor blocked）/ Step: first entry sensor blocked
    MUT_STEP_E2    : USINT := 2;        // 序列步：进入侧成对遮挡，屏蔽生效（Step: entry pair blocked, muting on）/ Step: entry pair blocked, muting on
    MUT_STEP_EXIT1 : USINT := 3;        // 序列步：首进入传感器清离（2 传感器退出段）/ Step: first entry sensor cleared (2-sensor exit)
    MUT_STEP_X1    : USINT := 4;        // 序列步：离开侧首传感器遮挡（4 传感器）/ Step: first exit sensor blocked (4-sensor)
    MUT_STEP_X2    : USINT := 5;        // 序列步：离开侧成对遮挡（4 传感器）/ Step: exit pair blocked (4-sensor)
    MUT_STEP_CL1   : USINT := 6;        // 序列步：离开侧首传感器清离（4 传感器退出段）/ Step: first exit sensor cleared (4-sensor exit)
END_VAR

METHOD CmdOverride : BOOL
VAR_INPUT
END_VAR
IF _bFaultLatch OR (_eState = E_DL_CurtainState.eFault) THEN
    CmdOverride := FALSE;         // 故障态拒绝（Rejected in fault）
ELSIF _bAnyMutBlocked THEN
    _bPendOverride := TRUE;       // 登记请求，主体编排消化（Register request, consumed by body）
    CmdOverride := TRUE;          // 受理成功（Accepted）
ELSE
    CmdOverride := FALSE;         // 无遮挡拒绝（Rejected with nothing blocked）
END_IF

(*------------------------------------------------------------------------------
 * 方法: CmdAck —— 屏蔽/故障确认复位：中止当前屏蔽序列回评估态（非故障态）。
 *      Method CmdAck - aborts the current muting sequence back to evaluation.
 *------------------------------------------------------------------------------*)
    END_METHOD

METHOD CmdAck : BOOL
VAR_INPUT
END_VAR
IF _bFaultLatch OR (_eState = E_DL_CurtainState.eFault) THEN
    CmdAck := FALSE;              // 故障态走 CmdReset（Fault goes through CmdReset）
ELSIF _bMutingAct OR _bOverrideAct THEN
    _bPendAck := TRUE;            // 登记确认请求（Register ack request）
    CmdAck := TRUE;               // 受理成功（Accepted）
ELSE
    CmdAck := FALSE;              // 无屏蔽活动可确认（Nothing to acknowledge）
END_IF

(*------------------------------------------------------------------------------
 * 方法: CmdReset —— 复位故障与重启联锁：仅故障态受理（接口方法拒绝语义）。
 *      Method CmdReset - reset fault and interlock, accepted only in fault.
 *------------------------------------------------------------------------------*)
    END_METHOD

METHOD CmdReset : BOOL
VAR_INPUT
END_VAR
IF _bFaultLatch OR (_eState = E_DL_CurtainState.eFault) THEN
    _bPendReset := TRUE;          // 登记复位请求（Register reset request）
    CmdReset := TRUE;             // 可复位（Resettable）
ELSE
    CmdReset := FALSE;            // 无故障可复位（Nothing to reset）
END_IF

(*------------------------------------------------------------------------------
 * 属性: eState（GET）—— 当前光幕状态只读视图。
 *      Property eState (GET) - read-only curtain state view.
 *------------------------------------------------------------------------------*)
    END_METHOD

// ============================================================================
// 段 1｜实例无条件周期刷新（R7/0.5：严禁置于 IF/CASE 分支内）
//      Unconditional per-cycle refresh of all instances (R7/0.5)
//      屏蔽灯闪烁用 TON 振荡器（IN := NOT Q 重触发）生成方波：Q 每 250MS 翻
//      转，override 态取 Q 作闪烁源；方波生成不适用 R14 断输入一拍规则（变
//      相位由振荡器自身承担），注释说明。
//      Lamp blink via a TON oscillator (IN := NOT Q): Q toggles every 250 MS;
//      the R14 one-scan-off rule does not apply to square-wave generation.
// ============================================================================
_fbTrigReset(CLK := bReset);
_fbTonDisc(IN := (bOssd1 <> bOssd2), PT := _tDiscEff);                    // OSSD 容差窗（OSSD discrepancy window）
_fbTonMutTo(IN := (_nMutStep > MUT_STEP_IDLE) AND (NOT _bFaultLatch), PT := _tMutToEff); // 屏蔽总时长（Muting total time）
_fbTonOvrMax(IN := _bOverrideAct, PT := _tOvrMaxEff);                     // override 硬帽（Override hard cap）
_fbTonBlink(IN := (NOT _fbTonBlink.Q), PT := DL_BLINK_HALF);              // 闪烁振荡器（Blink oscillator）

// ============================================================================
// 段 2｜参数钳位 + 信息级码预清零 + 复位路径（R15）
//      Parameter clamps + info preset + reset path (R15)
// ============================================================================
_uInfoCode := 0;                  // 信息级瞬时型每拍重算（Transient info recomputed each scan）
IF tMutingTimeout < DL_MUTTO_MIN THEN
    _tMutToEff := DL_MUTTO_MIN;   // 超时下限钳位（Timeout lower clamp）
ELSIF tMutingTimeout > DL_MUTTO_MAX THEN
    _tMutToEff := DL_MUTTO_MAX;   // 超时上限钳位（Timeout upper clamp）
ELSE
    _tMutToEff := tMutingTimeout; // 合法直通（Valid pass-through）
END_IF
IF tDiscrepancy < DL_DISC_MIN THEN
    _tDiscEff := DL_DISC_MIN;     // 容差窗下限钳位（Discrepancy lower clamp）
ELSIF tDiscrepancy > DL_DISC_MAX THEN
    _tDiscEff := DL_DISC_MAX;     // 容差窗上限钳位（Discrepancy upper clamp）
ELSE
    _tDiscEff := tDiscrepancy;    // 合法直通（Valid pass-through）
END_IF
IF tOverrideMax < DL_OVR_MIN THEN
    _tOvrMaxEff := DL_OVR_MIN;    // 硬帽下限钳位（Cap lower clamp）
ELSIF tOverrideMax > DL_OVR_MAX THEN
    _tOvrMaxEff := DL_OVR_MAX;    // 硬帽上限钳位（Cap upper clamp）
ELSE
    _tOvrMaxEff := tOverrideMax;  // 合法直通（Valid pass-through）
END_IF

IF _fbTrigReset.Q OR _bPendReset THEN
    _bPendReset := FALSE;         // 消费方法复位请求（Consume method reset）
    IF NOT _fbTonDisc.Q THEN      // 复位联锁：OSSD 不一致故障源已消失才解除（Restart interlock: source gone）
        _bFaultLatch := FALSE;    // 故障锁存解除（Fault latch released）
        _uErrorIdInt := 16#0000_0000; // 故障码清零（Fault code cleared）
        _nMutStep := MUT_STEP_IDLE;   // 序列步归零（Sequence step reset）
    END_IF
END_IF

// ============================================================================
// 段 3｜故障全局监视（优先级最高）：OSSD 双通道不一致 / 屏蔽超时
//      Global fault monitors: OSSD discrepancy / muting timeout
// ============================================================================
IF _fbTonDisc.Q THEN
    _bFaultLatch := TRUE;         // OSSD 双通道不一致锁存（OSSD discrepancy latch）
    _uErrorIdInt := 16#0003_02A2; // 0003_02A2 OSSD 双通道不一致【故障级】/ OSSD channel discrepancy, fault level
ELSIF _fbTonMutTo.Q THEN
    _bFaultLatch := TRUE;         // 屏蔽总时长超时锁存（Muting timeout latch）
    _uErrorIdInt := 16#0003_02A1; // 0003_02A1 屏蔽超时【故障级】/ Muting timeout, fault level
END_IF
IF _bFaultLatch THEN
    _nMutStep := MUT_STEP_IDLE;   // 故障即退出屏蔽序列（Fault exits the sequence）
END_IF

// ============================================================================
// 段 4｜传感器方向映射 + 屏蔽序列步进机 + override 编排（无故障时执行）
//      Sensor direction mapping + muting step machine + override orchestration
// ============================================================================
_bAnyMutBlocked := bMutSens1 OR bMutSens2 OR bMutSens3 OR bMutSens4; // 任一屏蔽传感器遮挡（Any sensor blocked）

IF NOT _bFaultLatch THEN
    // —— 方法确认消费：中止当前屏蔽/override 序列回评估态 ——
    IF _bPendAck THEN
        _bPendAck := FALSE;           // 消费方法确认请求（Consume method ack）
        _nMutStep := MUT_STEP_IDLE;   // 屏蔽序列中止（Sequence aborted）
        _bOverrideAct := FALSE;       // override 中止（Override aborted）
    END_IF

    // —— 方向映射（偏离②：首遮挡传感器判向）——
    IF bFourSensorMode THEN
        IF NOT _bMutRev THEN
            _bE1 := bMutSens1;        // 正向进入侧 1 = M1（Fwd entry 1 = M1）
            _bE2 := bMutSens2;        // 正向进入侧 2 = M2（Fwd entry 2 = M2）
            _bX1 := bMutSens3;        // 正向离开侧 1 = M3（Fwd exit 1 = M3）
            _bX2 := bMutSens4;        // 正向离开侧 2 = M4（Fwd exit 2 = M4）
        ELSE
            _bE1 := bMutSens4;        // 反向进入侧 1 = M4（Rev entry 1 = M4）
            _bE2 := bMutSens3;        // 反向进入侧 2 = M3（Rev entry 2 = M3）
            _bX1 := bMutSens2;        // 反向离开侧 1 = M2（Rev exit 1 = M2）
            _bX2 := bMutSens1;        // 反向离开侧 2 = M1（Rev exit 2 = M1）
        END_IF
    ELSE
        IF NOT _bMutRev THEN
            _bE1 := bMutSens1;        // 正向进入侧 1 = M1（Fwd entry 1 = M1）
            _bE2 := bMutSens2;        // 正向进入侧 2 = M2（Fwd entry 2 = M2）
        ELSE
            _bE1 := bMutSens2;        // 反向进入侧 1 = M2（Rev entry 1 = M2）
            _bE2 := bMutSens1;        // 反向进入侧 2 = M1（Rev entry 2 = M1）
        END_IF
        _bX1 := _bE1;                 // 2 传感器模式：离开侧=同对清离（Exit = clearing of the same pair）
        _bX2 := _bE2;
    END_IF

    // —— 屏蔽序列步进机（电平条件级联，序列错乱即故障退出）——
    //     Muting sequence step machine (level-condition cascade, any deviation faults out)
    IF NOT bEnableMuting THEN
        _nMutStep := MUT_STEP_IDLE;   // 总使能切断：序列强制空闲（Master disable forces idle）
    ELSE
        CASE _nMutStep OF
            MUT_STEP_IDLE: // 空闲：等待首传感器遮挡判向
                IF _bE1 AND (NOT _bE2) AND (NOT _bX1) AND (NOT _bX2) THEN
                    _nMutStep := MUT_STEP_E1; // 首进入传感器遮挡（First entry sensor blocked）
                ELSIF ((NOT bFourSensorMode) AND _bE2 AND (NOT _bE1))
                   OR (bFourSensorMode AND _bX2 AND (NOT _bE1) AND (NOT _bE2) AND (NOT _bX1)) THEN
                    _bMutRev := NOT _bMutRev; // 次序第二传感器先遮挡：判反向（v1.0.1 修复：原条件 2 传感器
                                              // 模式与正向 IF 恒等矛盾成死代码、4 传感器模式误查 M3，
                                              // 按偏离②语义 M2/M4 先遮挡=反向）/ Second-in-order blocked
                                              // first: reverse (v1.0.1 fix per deviation note ②)
                    _nMutStep := MUT_STEP_E1; // 反向序列启动（Reverse sequence starts）
                END_IF

            MUT_STEP_E1: // 首进入传感器已遮挡：等第二进入传感器
                IF _bE1 AND _bE2 THEN
                    _nMutStep := MUT_STEP_E2; // 进入侧成对遮挡，屏蔽生效（Entry pair blocked, muting on）
                ELSIF NOT _bE1 THEN
                    _bFaultLatch := TRUE;     // 首传感器提前清离：序列错乱（First sensor cleared early: sequence error）
                    _uErrorIdInt := 16#0003_02A0; // 0003_02A0 屏蔽传感器序列错误【故障级】/ Muting sequence error, fault level
                    _nMutStep := MUT_STEP_IDLE;
                END_IF

            MUT_STEP_E2: // 屏蔽生效：2 传感器等首清离 / 4 传感器等离开侧首遮挡
                IF bFourSensorMode THEN
                    IF _bX1 THEN
                        _nMutStep := MUT_STEP_X1; // 离开侧首传感器遮挡（First exit sensor blocked）
                    ELSIF (NOT _bE1) OR (NOT _bE2) THEN
                        _nMutStep := MUT_STEP_IDLE; // 物未达离开侧即全清：屏蔽正常收尾（Cleared before exit pair: normal end）
                    ELSIF _bX2 THEN
                        _bFaultLatch := TRUE;     // 离开侧第二传感器先遮挡：序列错乱（Exit second first: sequence error）
                        _uErrorIdInt := 16#0003_02A0;
                        _nMutStep := MUT_STEP_IDLE;
                    END_IF
                ELSE
                    IF (NOT _bE1) AND _bE2 THEN
                        _nMutStep := MUT_STEP_EXIT1; // 首进入传感器清离（First entry sensor cleared）
                    ELSIF (NOT _bE2) AND _bE1 THEN
                        _bFaultLatch := TRUE;        // 第二传感器先清离：序列错乱（Second cleared first: sequence error）
                        _uErrorIdInt := 16#0003_02A0;
                        _nMutStep := MUT_STEP_IDLE;
                    ELSIF (NOT _bE1) AND (NOT _bE2) THEN
                        _nMutStep := MUT_STEP_IDLE;  // 双清离：物体回退/中断恢复，序列中止回评估态（v1.0.1 修复：
                                                     // 原无分支滞留 E2 依赖屏蔽超时误报故障）/ Both cleared:
                                                     // abort back to evaluation (v1.0.1 fix)
                    END_IF
                END_IF

            MUT_STEP_EXIT1: // 2 传感器退出段：等第二传感器清离
                IF (NOT _bE1) AND (NOT _bE2) THEN
                    _nMutStep := MUT_STEP_IDLE;   // 序列完成（Sequence complete）
                ELSIF _bE1 AND _bE2 THEN
                    _nMutStep := MUT_STEP_E2;     // 新物体衔接进入：回屏蔽段（Back-to-back object: back to muting）
                END_IF

            MUT_STEP_X1: // 4 传感器：离开侧首遮挡，等成对
                IF _bX1 AND _bX2 THEN
                    _nMutStep := MUT_STEP_X2;     // 离开侧成对遮挡（Exit pair blocked）
                ELSIF NOT _bX1 THEN
                    _bFaultLatch := TRUE;         // 离开首传感器提前清离：序列错乱（Exit first cleared early: error）
                    _uErrorIdInt := 16#0003_02A0;
                    _nMutStep := MUT_STEP_IDLE;
                END_IF

            MUT_STEP_X2: // 4 传感器：离开侧成对，等首清离
                IF (NOT _bX1) AND _bX2 THEN
                    _nMutStep := MUT_STEP_CL1;    // 离开首传感器清离（Exit first cleared）
                ELSIF (NOT _bX2) AND _bX1 THEN
                    _bFaultLatch := TRUE;         // 离开第二传感器先清离：序列错乱（Exit second cleared first: error）
                    _uErrorIdInt := 16#0003_02A0;
                    _nMutStep := MUT_STEP_IDLE;
                END_IF

            MUT_STEP_CL1: // 4 传感器退出段：等第二传感器清离
                IF (NOT _bX1) AND (NOT _bX2) THEN
                    _nMutStep := MUT_STEP_IDLE;   // 序列完成（Sequence complete）
                ELSIF _bX1 AND _bX2 THEN
                    _nMutStep := MUT_STEP_X2;     // 新物体衔接：回成对段（Back-to-back: back to pair state）
                END_IF

            ELSE
                _nMutStep := MUT_STEP_IDLE;       // 步号域外兜底：强制空闲（Out-of-domain step: force idle）
        END_CASE
    END_IF

    // —— override 编排：准入硬约束（钥匙/方法请求 AND 至少一传感器遮挡）——
    //     Override orchestration: admission hard constraint
    IF _bOverrideAct THEN
        IF (NOT bOverrideKey) AND (NOT _bPendOverride) THEN
            _bOverrideAct := FALSE;       // 请求撤销退出（Request dropped: exit override）
        ELSIF _fbTonOvrMax.Q THEN
            _bOverrideAct := FALSE;       // 硬帽到期退出（Hard cap expired: exit override）
            _uInfoCode := 16#0003_0118;   // 0003_0118 override 硬帽到期退出【信息级】/ Override cap exit, info level
        END_IF
    ELSE
        IF (bOverrideKey OR _bPendOverride) AND _bAnyMutBlocked AND (NOT _bFaultLatch) THEN
            _bOverrideAct := TRUE;        // 准入成立进入 override（Admission granted, enter override）
        ELSIF (bOverrideKey OR _bPendOverride) AND (NOT _bAnyMutBlocked) THEN
            _uInfoCode := 16#0003_0122;   // 0003_0122 override 准入拒绝（无遮挡）【信息级】/ Override denied (nothing blocked), info level
        END_IF
        _bPendOverride := FALSE;          // 方法请求消费（Method request consumed）
    END_IF
END_IF

_bMutingAct := (_nMutStep >= MUT_STEP_E2) AND (NOT _bFaultLatch); // 屏蔽生效派生（Muting-active derived form）

// ============================================================================
// 段 5｜状态映像（IF 派生链含 ELSE 兜底）+ 输出推导 + bSafeStop 出口断言
//      State image (IF derivation chain with ELSE) + outputs + bSafeStop assertion
// ============================================================================
IF _bFaultLatch THEN
    _eState := E_DL_CurtainState.eFault;            // 故障锁存映像（Fault image）
ELSIF _bOverrideAct THEN
    _eState := E_DL_CurtainState.eOverride;         // 滞留清除映像（Override image）
ELSIF _bMutingAct THEN
    _eState := E_DL_CurtainState.eMuting;           // 屏蔽进行中映像（Muting image）
ELSIF NOT (bOssd1 AND bOssd2) THEN
    _eState := E_DL_CurtainState.eBlocked;          // 遮挡未屏蔽映像（Blocked image）
ELSE
    _eState := E_DL_CurtainState.eClear;            // 通光兜底映像（Clear fallback image）
END_IF

// bSafeStop 不在此处赋值：其为接口属性，由 PROPERTY bSafeStop（GET）以出口
// 断言式承载（R22）；此处仅推导非接口输出 bMutingLamp。
// bSafeStop is not written here: as an interface attribute it is carried by the
// PROPERTY getter with exit assertion (R22); only bMutingLamp is derived here.
bMutingLamp := _bMutingAct OR (_bOverrideAct AND _fbTonBlink.Q); // 屏蔽灯：屏蔽常亮/override 闪烁（Lamp: steady/blink）

(*------------------------------------------------------------------------------
 * 方法: CmdOverride —— 滞留物清除请求：至少一个屏蔽传感器仍遮挡才受理。
 *      Method CmdOverride - override accepted only with a muting sensor blocked.
 *------------------------------------------------------------------------------*)

PROPERTY eState : E_DL_CurtainState
eState := _eState;                // 返回派生状态（Return derived state）

(*------------------------------------------------------------------------------
 * 属性: bClear（GET）—— 光幕通光（OSSD 双通道全通光）。
 *      Property bClear (GET) - curtain clear (both OSSD channels clear).
 *------------------------------------------------------------------------------*)
PROPERTY bClear : BOOL
bClear := bOssd1 AND bOssd2;      // 双通道通光派生式（Both-channel clear derived form）

(*------------------------------------------------------------------------------
 * 属性: bMutingActive（GET）—— 屏蔽进行中。
 *      Property bMutingActive (GET) - muting active.
 *------------------------------------------------------------------------------*)
PROPERTY bMutingActive : BOOL
bMutingActive := _bMutingAct;     // 返回屏蔽派生标志（Return muting derived flag）

(*------------------------------------------------------------------------------
 * 属性: bOverrideActive（GET）—— 滞留清除进行中。
 *      Property bOverrideActive (GET) - override active.
 *------------------------------------------------------------------------------*)
PROPERTY bOverrideActive : BOOL
bOverrideActive := _bOverrideAct; // 返回 override 标志（Return override flag）

(*------------------------------------------------------------------------------
 * 属性: bSafeStop（GET）—— 应停机输出（核心安全镜像位，屏蔽/override 态断
 *         言恒 FALSE，永不因屏蔽置假）。
 *      Property bSafeStop (GET) - safe-stop mirror, asserted FALSE when muting/override.
 *------------------------------------------------------------------------------*)
PROPERTY bSafeStop : BOOL
bSafeStop := (NOT (bOssd1 AND bOssd2)) AND (NOT _bMutingAct)
          AND (NOT _bOverrideAct) AND (NOT _bFaultLatch); // 出口断言式派生（Exit-assertion derived form）

(*------------------------------------------------------------------------------
 * 属性: bFault（GET）—— 故障锁存指示（信息级码不置本位，0.2 公约）。
 *      Property bFault (GET) - fault latch indicator, info codes excluded.
 *------------------------------------------------------------------------------*)
PROPERTY bFault : BOOL
bFault := _bFaultLatch OR (_eState = E_DL_CurtainState.eFault); // 显式排除信息级派生式（Derived form excluding info codes）

(*------------------------------------------------------------------------------
 * 属性: uErrorId（GET）—— 末次故障码（故障级优先，无故障时透出本拍信息级
 *         码，0.2/0.15 公约）。
 *      Property uErrorId (GET) - last error code (fault priority, info shown otherwise).
 *------------------------------------------------------------------------------*)
PROPERTY uErrorId : UDINT
IF (_uErrorIdInt <> 0) OR (_eState = E_DL_CurtainState.eFault) THEN
    uErrorId := _uErrorIdInt;     // 故障级码优先透出（Fault-level priority）
ELSE
    uErrorId := _uInfoCode;       // 无故障时透出本拍信息级码（Transient info code）
END_IF
END_FUNCTION_BLOCK
